(* IEC 61131-3 sources: plcassist-cli/packages/volt-lsp-iec/test-corpus/bakon-nano/Device/Plc Logic/Application/POUs/Calculations (part 2) *)

(* ---- Calc_Hor.fun ---- *)
function Calc_Hor : bool
VAR
	nNrOfLines: INT;
	rLengthOfLine: REAL;
	nNumberOfCutsPerLine: INT;
	nCnt_pos: INT;
	nCnt_line: INT;
	nCnt_Push: INT;
	bToggle: BOOL;
	//nFirstPos: INT;
	//nFirstWastePos: INT;
	rLast_Y_Pos	:REAL;
	rSizeTrimRear	:REAL;
	rSizeTrimFront	:REAL;
	rSizeTrimRight	:REAL;
	rSizeTrimLeft	:REAL;

	//CorrectOvershootHor1a	: CorrectOvershootHor;
	//CorrectOvershootHor1b	: CorrectOvershootHor;
	//CorrectOvershootHor2	: CorrectOvershootHor;
	//CorrectOvershootHor3	: CorrectOvershootHor;
	//CorrectOvershootHor4	: CorrectOvershootHor;
	//CorrectOvershootHor5	: CorrectOvershootHor;
	//CorrectOvershootHor6	: CorrectOvershootHor;
	//CorrectOvershootHor7	: CorrectOvershootHor;
	rMaxTraySize: REAL;
	rMinTraySize: REAL;
	rProdLength_InY: REAL;
	rProdLength_InX: REAL;
	rMmPerCut :REAL;
	rCenterPointKnifeInverted: REAL;
	rSizeOfKnife: REAL;
	//rStartPointTray_Y: REAL;
	rMinimumTrayTrimSize: REAL;
	rNrOfLines 	:REAL;
	rWasteExtra	:REAL;
	rIcedOffset	:REAL;

	rCenterPointKnife: REAL;
	rMinimumSlabTrimSize: REAL;
	nPartsY: INT;

	FirstPoint					: Gonio_Point;
	CopyPoint					: Gonio_Point;

	rFirstYPosition : REAL;
	overshootSettings 			: Gonio_Settings;
	nFirstPosFirstTray 		:INT;
	nFirstWastePosFirstTray :INT;
	nLastPosFirstTray		: INT;
	nLastWastePosFirstTray	: int;
END_VAR

(* Calc_Hor, (mes 0 graden *)

(************************************************************************************************************************************
 * HISTORY
 ************************************************************************************************************************************
 * Update 		: 0.1
 * Author 		: K. Kole
 * Changes	: Tray square, 	calculation for rSizeTrimRight and rSizeTrimLeft changed
 * Update 		: 0.2
 * Author 		: K. Kole
 * Changes	: Tray square, 	calculation for rSizeTrimRear and rSizeTrimFront changed
 ************************************************************************************************************************************)
Calc_Hor := FALSE;
bToggle	:= FALSE;
//nFirstPos := g_sCuttingPositionsInfo.index;
//nFirstWastePos := g_sWastePositionsInfo.index ;

nFirstPosFirstTray 				:= g_sCuttingPositionsInfo.index;
nFirstWastePosFirstTray 		:= g_sWastePositionsInfo.index;

rSizeOfKnife					:= g_HMI_MCH_Parameters.rSizeOfKnife;
rCenterPointKnife				:= rSizeOfKnife/2;
rCenterPointKnifeInverted	:= rSizeOfKnife/2;

overshootSettings.knifeAxis		:= rCenterPointKnife;
overshootSettings.knifeLength	:= rSizeOfKnife;
overshootSettings.precision		:= 0.1;

(**********************************************************************************************************************************)
(* Tray square *)(*AC 23-10-2012 Also Tray Triangle*)
(**********************************************************************************************************************************)
IF		((g_HMI_RCP_Parameters.nProductType = Prod_Tray_Rectangle_1x1)
	OR	(g_HMI_RCP_Parameters.nProductType = Prod_Tray_Rectangle_1x2)
	OR	(g_HMI_RCP_Parameters.nProductType = Prod_Tray_Rectangle_1x4)
	OR 	(g_HMI_RCP_Parameters.nProductType = Prod_Tray_Rectangle_2x1))
THEN

	(* Determine type of tray *)
	IF  (g_HMI_RCP_Parameters.nProductType = Prod_Tray_Rectangle_1x1) THEN
		rProdLength_InY	:= g_HMI_MCH_Parameters.rProdLengthTrayLarge_InY;
		rProdLength_InX	:= g_HMI_MCH_Parameters.rProdLengthTrayLarge_InX;
		rMinimumTrayTrimSize :=	g_HMI_MCH_Parameters.rMinimumTrimSizeTrayLarge;
		FirstPoint.X := g_HMI_MCH_Parameters.rStartPointTrayLarge_X;
		FirstPoint.Y := g_HMI_MCH_Parameters.rStartPointTrayLarge_Y;
	ELSIF	(g_HMI_RCP_Parameters.nProductType = Prod_Tray_Rectangle_1x2)
	THEN
		rProdLength_InY	:= g_HMI_MCH_Parameters.rProdLengthTraySmall_InY;
		rProdLength_InX	:= g_HMI_MCH_Parameters.rProdLengthTraySmall_InX;
		rMinimumTrayTrimSize :=	g_HMI_MCH_Parameters.rMinimumTrimSizeTraySmall;
		FirstPoint.X  := g_HMI_MCH_Parameters.rStartPointTraySmall_X;
		FirstPoint.Y  := g_HMI_MCH_Parameters.rStartPointTraySmall1_Y;	(* Startpoint for first small tray *)
	ELSIF	(g_HMI_RCP_Parameters.nProductType = Prod_Tray_Rectangle_1x4)
	THEN
		rProdLength_InY	:= g_HMI_MCH_Parameters.rProdLengthTrayTriple_InY;
		rProdLength_InX	:= g_HMI_MCH_Parameters.rProdLengthTrayTriple_InX;
		rMinimumTrayTrimSize :=	g_HMI_MCH_Parameters.rMinimumTrimSizeTrayTriple;
		FirstPoint.X  := g_HMI_MCH_Parameters.rStartPointTrayTriple_X;
		FirstPoint.Y  := g_HMI_MCH_Parameters.rStartPointTrayTriple1_Y;	(* Startpoint for first small tray *)
	ELSIF	(g_HMI_RCP_Parameters.nProductType = Prod_Tray_Rectangle_2x1)
	THEN
		rProdLength_InY	:= g_HMI_MCH_Parameters.rProdLengthTrayDouble_InY;
		rProdLength_InX	:= g_HMI_MCH_Parameters.rProdLengthTrayDouble_InX;
		rMinimumTrayTrimSize :=	g_HMI_MCH_Parameters.rMinimumTrimSizeTrayDouble;
		FirstPoint.X  := g_HMI_MCH_Parameters.rStartPointTrayDouble1_X;
		FirstPoint.Y  := g_HMI_MCH_Parameters.rStartPointTrayDouble_Y;	(* Startpoint for first small tray *)
	END_IF

	IF g_HMI_RCP_Parameters.bTrianglesInTray AND g_HMI_RCP_Parameters.bUseRectanglesInEight THEN (*AC 04-07-2013: Uitbreiding 8 driehoeken uit stuk*)
		nPartsY := g_HMI_RCP_Parameters.nPartsY * 2;
	ELSE
		nPartsY := g_HMI_RCP_Parameters.nPartsY;
	END_IF

	IF g_HMI_RCP_Parameters.rSizeTrimFront <= 0			(* Wijziging 16 juli 2010 *)(*AC 28-11-12: Omgedraaid vanaf HMI INstellingen*)
	THEN
		rSizeTrimRear	:= 0;
	ELSE
		rSizeTrimRear 	:= MAX(rMinimumTrayTrimSize, g_HMI_RCP_Parameters.rSizeTrimFront); (*AC 28-11-12: Omgedraaid vanaf HMI INstellingen*)
	END_IF
	IF g_HMI_RCP_Parameters.rSizeTrimRear<= 0			(* Wijziging 16 juli 2010 *)(*AC 28-11-12: Omgedraaid vanaf HMI INstellingen*)
	THEN
		rSizeTrimFront	:= 0;
	ELSE
		rSizeTrimFront 	:= MAX(rMinimumTrayTrimSize, g_HMI_RCP_Parameters.rSizeTrimRear);(*AC 28-11-12: Omgedraaid vanaf HMI INstellingen*)
	END_IF
	rSizeTrimRight 	:= MAX(rMinimumTrayTrimSize, g_HMI_RCP_Parameters.rSizeTrimRight);
	rSizeTrimLeft 		:= MAX(rMinimumTrayTrimSize, g_HMI_RCP_Parameters.rSizeTrimLeft);

	(*Additional safety checks for trays*)
	rMaxTraySize := rProdLength_InX - (rMinimumTrayTrimSize * 2);
	IF			rMaxTraySize >= (g_HMI_MCH_Parameters.rSizeOfKnife)											(* Fixed mes past in het blik *)
	THEN
		rSizeOfKnife					:= g_HMI_MCH_Parameters.rSizeOfKnife;
		rCenterPointKnife				:= rSizeOfKnife/2;
		rCenterPointKnifeInverted	:= rSizeOfKnife/2;
		rMinTraySize					:= rProdLength_InX - (rSizeTrimRight + rSizeTrimLeft);
		IF rMinTraySize < rSizeOfKnife THEN
			rSizeTrimRight	:= rSizeTrimRight - (rSizeOfKnife - rMinTraySize);
			rSizeTrimRight 	:= MAX(rMinimumTrayTrimSize, rSizeTrimRight);								(* Check if new calculated trim is >= MinimumTrim *)
			rSizeTrimLeft	:= rProdLength_InX - rSizeOfKnife - rSizeTrimRight;
		END_IF
	ELSE																											(* Fixed mes past NIET in het blik *)
		g_sMACH.ERR.bTrayTooSmall := TRUE;
		RETURN;
	END_IF

	g_rDistanceBetweenCuts_InY:=	(rProdLength_InY - rSizeTrimRear - rSizeTrimFront) / INT_TO_REAL(nPartsY);(*g_HMI_RCP_Parameters.nPartsY);*)

	(* Determine number of lines *)
	IF g_bTrimRear AND g_bTrimFront
	THEN
		nNrOfLines	:= 1 + nPartsY;(*g_HMI_RCP_Parameters.nPartsY);*)(*AC 04-07-2013*)
	ELSIF g_bTrimRear AND NOT g_bTrimFront
	THEN
		nNrOfLines	:= nPartsY;(*g_HMI_RCP_Parameters.nPartsY);*)(*AC 04-07-2013*)
	ELSIF NOT g_bTrimRear AND g_bTrimFront
	THEN
		nNrOfLines	:= nPartsY;(*g_HMI_RCP_Parameters.nPartsY);*)(*AC 04-07-2013*)
	ELSIF NOT g_bTrimRear AND NOT g_bTrimFront
	THEN
		nNrOfLines	:=nPartsY - 1;(*g_HMI_RCP_Parameters.nPartsY);*)(*AC 04-07-2013*)
	END_IF

	(* Calculate number of cuts on the line *)
	rLengthOfLine := rProdLength_InX - rSizeTrimRight - rSizeTrimLeft;
	IF rLengthOfLine > rSizeOfKnife
	THEN
		nNumberOfCutsPerLine := TRUNC_INT(rLengthOfLine / rSizeOfKnife);
		IF nNumberOfCutsPerLine < (rLengthOfLine / rSizeOfKnife)
		THEN
			nNumberOfCutsPerLine := nNumberOfCutsPerLine + 1;
		END_IF
	ELSE
		nNumberOfCutsPerLine := 1;
	END_IF
	(*Calculation of covered distance per cut*)
	rMmPerCut := (rLengthOfLine - rSizeOfKnife)/(nNumberOfCutsPerLine -1);

	(* Calculate positions on first line *)
	overshootSettings.MarginXMin := FirstPoint.x + MAX(rMinimumTrayTrimSize-0.1,1);		(* Mechanical boundary *)
	overshootSettings.MarginXMax := FirstPoint.x + rProdLength_InX  - MAX(rMinimumTrayTrimSize-0.1,1);	(* Mechanical boundary *)
	overshootSettings.MarginYMin := FirstPoint.y + MAX(rMinimumTrayTrimSize-0.1,1);		(* Mechanical boundary *)
	overshootSettings.MarginYMax := FirstPoint.y + rProdLength_InY -  MAX(rMinimumTrayTrimSize-0.1,1);		(* Mechanical boundary *)

	overshootSettings.adjustXMax := FALSE;
	overshootSettings.adjustXMin := FALSE;
	overshootSettings.adjustYMax := FALSE;
	overshootSettings.adjustYMin := FALSE;

	IF g_bTrimRear
	THEN
		IF nNumberOfCutsPerLine = 1
		THEN
			IF NOT StorePos(I_rX:= 							Firstpoint.X + rSizeTrimRight + rCenterPointKnife,
							I_rY:=							(rFirstYPosition := Firstpoint.Y + rSizeTrimRear),
							I_rA:=							0,
							I_rK:=							0,
							I_bIsWaste :=					 (g_HMI_RCP_Parameters.bCutWasteFirst) ,
							I_sOvershootSettings := 		overshootSettings)
			THEN
								RETURN;
			END_IF
		ELSE
			FOR nCnt_pos:=1 TO (nNumberOfCutsPerLine - 1) DO
				IF NOT StorePos(I_rX:= 							FirstPoint.X + rSizeTrimRight + (nCnt_pos - 1) * rMmPerCut
																			 + rCenterPointKnife,
								I_rY:=							(rFirstYPosition := FirstPoint.Y + rSizeTrimRear),
								I_rA:=							0,
								I_rK:=							0,
								I_bIsWaste :=					 (g_HMI_RCP_Parameters.bCutWasteFirst) ,
								I_sOvershootSettings := 		overshootSettings)
				THEN
										RETURN;
				END_IF
			END_FOR
			(* Last position on the line *)
			IF NOT StorePos(I_rX:= 							Firstpoint.X + rProdLength_InX - rSizeTrimLeft - rCenterPointKnifeInverted,
							I_rY:=							Firstpoint.Y + rSizeTrimRear,
							I_rA:=							0,
							I_rK:=							0,
							I_bIsWaste :=					 (g_HMI_RCP_Parameters.bCutWasteFirst) ,
							I_sOvershootSettings := 		overshootSettings)
			THEN
								RETURN;
			END_IF

		END_IF
	ELSE (* No waste strip at the left *)
		IF nNrOfLines > 0	(* New 8 feb 2010: when only one piece and no trims *)
		THEN
			IF nNumberOfCutsPerLine = 1
			THEN
				IF NOT StorePos(I_rX:= 							Firstpoint.X + rSizeTrimRight + rCenterPointKnife,
								I_rY:=							(rFirstYPosition := Firstpoint.Y + rSizeTrimRear + g_rDistanceBetweenCuts_InY),
								I_rA:=							0,
								I_rK:=							0,
								I_bIsWaste :=					FALSE,
								I_sOvershootSettings := 		overshootSettings)
				THEN
										RETURN;
				END_IF

			ELSE
				FOR nCnt_pos:=1 TO (nNumberOfCutsPerLine - 1) DO
					IF NOT StorePos(I_rX:= 							Firstpoint.X + rSizeTrimRight + (nCnt_pos - 1) * rMmPerCut
																					 + rCenterPointKnife,
									I_rY:=							(rFirstYPosition := Firstpoint.Y + rSizeTrimRear + g_rDistanceBetweenCuts_InY),
									I_rA:=							0,
									I_rK:=							0,
									I_bIsWaste :=					FALSE,
									I_sOvershootSettings := 		overshootSettings)
					THEN
												RETURN;
					END_IF

				END_FOR
				(* Last position on the line *)
				IF NOT StorePos(I_rX:= 							Firstpoint.X + rProdLength_InX - rSizeTrimLeft - rCenterPointKnifeInverted,
								I_rY:=							Firstpoint.Y + rSizeTrimRear + g_rDistanceBetweenCuts_InY,
								I_rA:=							0,
								I_rK:=							0,
								I_bIsWaste :=					FALSE,
								I_sOvershootSettings := 		overshootSettings)
				THEN
										RETURN;
				END_IF

			END_IF
		END_IF
	END_IF

	(* Fill in all other positions on the rest of the lines *)

	FOR nCnt_line := 2 TO (nNrOfLines) BY 1 DO
		IF nNumberOfCutsPerLine = 1
		THEN
			IF NOT StorePos(I_rX:= 							Firstpoint.X + rSizeTrimRight + rCenterPointKnife,
							I_rY:=							rFirstYPosition + (nCnt_line-1) * g_rDistanceBetweenCuts_InY,
							I_rA:=							0,
							I_rK:=							0,
							I_bIsWaste :=					 (g_HMI_RCP_Parameters.bCutWasteFirst AND g_bTrimFront AND nCnt_Line = nNrOfLines) ,
							I_sOvershootSettings := 		overshootSettings)
			THEN
								RETURN;
			END_IF

		ELSE
			IF bToggle (* from front to rear *)
			THEN
				FOR nCnt_pos:=1 TO (nNumberOfCutsPerLine - 1) DO
					IF NOT StorePos(I_rX:= 							Firstpoint.X + rSizeTrimRight + rCenterPointKnife
														                                                   + (nCnt_pos - 1) * rMmPerCut ,
									I_rY:=							rFirstYPosition + (nCnt_line-1) * g_rDistanceBetweenCuts_InY,
									I_rA:=							0,
									I_rK:=							0,
									I_bIsWaste :=					 (g_HMI_RCP_Parameters.bCutWasteFirst AND g_bTrimFront AND nCnt_Line = nNrOfLines) ,
									I_sOvershootSettings := 		overshootSettings)
					THEN
												RETURN;
					END_IF

				END_FOR
				(* Last position on the line *)
				IF NOT StorePos(I_rX:= 							Firstpoint.X + rProdLength_InX - rSizeTrimLeft - rCenterPointKnifeInverted,
								I_rY:=							rFirstYPosition + (nCnt_line-1) * g_rDistanceBetweenCuts_InY,
								I_rA:=							0,
								I_rK:=							0,
								I_bIsWaste :=					 (g_HMI_RCP_Parameters.bCutWasteFirst AND g_bTrimFront AND nCnt_Line = nNrOfLines) ,
								I_sOvershootSettings := 		overshootSettings)
				THEN
										RETURN;
				END_IF

			ELSE (* toggle, ie from rear to front *)
				FOR nCnt_pos:=1 TO (nNumberOfCutsPerLine - 1) DO
					IF NOT StorePos(I_rX:= 							Firstpoint.X + rProdLength_InX - rSizeTrimLeft - rCenterPointKnifeInverted
																					- (nCnt_pos -1) * rMmPerCut,
									I_rY:=							rFirstYPosition + (nCnt_line-1) * g_rDistanceBetweenCuts_InY,
									I_rA:=							0,
									I_rK:=							0,
									I_bIsWaste :=					 (g_HMI_RCP_Parameters.bCutWasteFirst AND g_bTrimFront AND nCnt_Line = nNrOfLines) ,
									I_sOvershootSettings := 		overshootSettings)
					THEN
												RETURN;
					END_IF

				END_FOR
				(* Last position on the line *)
				IF NOT StorePos(I_rX:= 							FirstPoint.X + rSizeTrimRight + rCenterPointKnife,
								I_rY:=							rFirstYPosition + (nCnt_line-1) * g_rDistanceBetweenCuts_InY,
								I_rA:=							0,
								I_rK:=							0,
								I_bIsWaste :=					 (g_HMI_RCP_Parameters.bCutWasteFirst AND g_bTrimFront AND nCnt_Line = nNrOfLines) ,
								I_sOvershootSettings := 		overshootSettings)
				THEN
										RETURN;
				END_IF

			END_IF
			bToggle := NOT bToggle;
		END_IF
	END_FOR

	nLastPosFirstTray		:= g_sCuttingPositionsInfo.index-1;
	nLastWastePosFirstTray	:= g_sWastePositionsInfo.index-1;

	(* Double the positions for the second tray if small trays is selected *)
	IF	g_HMI_RCP_Parameters.nProductType = Prod_Tray_Rectangle_1x2
	THEN

		CopyPoint.X := FirstPoint.X;
		CopyPoint.Y := g_HMI_MCH_Parameters.rStartPointTraySmall2_Y;

		overshootSettings.MarginXMin := CopyPoint.X + MAX(rMinimumTrayTrimSize-0.1,1);		(* Mechanical boundary *)
		overshootSettings.MarginXMax := CopyPoint.X + rProdLength_InX  - MAX(rMinimumTrayTrimSize-0.1,1);	(* Mechanical boundary *)
		overshootSettings.MarginYMin := CopyPoint.Y + MAX(rMinimumTrayTrimSize-0.1,1);		(* Mechanical boundary *)
		overshootSettings.MarginYMax := CopyPoint.Y + rProdLength_InY -  MAX(rMinimumTrayTrimSize-0.1,1);		(* Mechanical boundary *)

		IF nFirstPosFirstTray <= nLastPosFirstTray THEN
			IF NOT Calc_CopyCutsWithOffset(
				I_firstIndex				:= nFirstPosFirstTray,
				I_lastIndex					:= nLastPosFirstTray,
				I_dX 						:= CopyPoint.X - FirstPoint.X,
				I_dY 						:= CopyPoint.Y - FirstPoint.Y,
				I_overshootSettings 		:= overshootSettings,
				I_dataArray 				:= ADR(g_aCuttingPositions),
				I_bReverseOrder				:= (nNrOfLines MOD 2)>0,
				IQ_dataArrayInfo 			:= g_sCuttingPositionsInfo)
			THEN
								RETURN;
			END_IF
		END_IF

		IF nFirstWastePosFirstTray <= nLastWastePosFirstTray THEN
			IF NOT Calc_CopyCutsWithOffset(
				I_firstIndex				:= nFirstWastePosFirstTray,
				I_lastIndex					:= nLastWastePosFirstTray,
				I_dX 						:= CopyPoint.X - FirstPoint.X,
				I_dY 						:= CopyPoint.Y - FirstPoint.Y,
				I_overshootSettings 		:= overshootSettings,
				I_dataArray 				:= ADR(g_aWastePositions),
				I_bReverseOrder				:= (nNrOfLines MOD 2)>0,
				IQ_dataArrayInfo 			:= g_sWastePositionsInfo)
			THEN
								RETURN;
			END_IF
		END_IF
	END_IF

	(* Triple the positions for the second and third tray if triple trays is selected *)
	IF	g_HMI_RCP_Parameters.nProductType = Prod_Tray_Rectangle_1x4
	THEN

		CopyPoint.X := FirstPoint.X;
		CopyPoint.Y := g_HMI_MCH_Parameters.rStartPointTrayTriple2_Y;

		overshootSettings.MarginXMin := CopyPoint.X + MAX(rMinimumTrayTrimSize-0.1,1);		(* Mechanical boundary *)
		overshootSettings.MarginXMax := CopyPoint.X + rProdLength_InX  - MAX(rMinimumTrayTrimSize-0.1,1);	(* Mechanical boundary *)
		overshootSettings.MarginYMin := CopyPoint.Y + MAX(rMinimumTrayTrimSize-0.1,1);		(* Mechanical boundary *)
		overshootSettings.MarginYMax := CopyPoint.Y + rProdLength_InY -  MAX(rMinimumTrayTrimSize-0.1,1);		(* Mechanical boundary *)

		IF nFirstPosFirstTray <= nLastPosFirstTray THEN
			IF NOT Calc_CopyCutsWithOffset(
				I_firstIndex				:= nFirstPosFirstTray,
				I_lastIndex					:= nLastPosFirstTray,
				I_dX 						:= CopyPoint.X - FirstPoint.X,
				I_dY 						:= CopyPoint.Y - FirstPoint.Y,
				I_overshootSettings 		:= overshootSettings,
				I_dataArray 				:= ADR(g_aCuttingPositions),
				I_bReverseOrder				:= (nNrOfLines MOD 2)>0,
				IQ_dataArrayInfo 			:= g_sCuttingPositionsInfo)
			THEN
								RETURN;
			END_IF
		END_IF

		IF nFirstWastePosFirstTray <= nLastWastePosFirstTray THEN
			IF NOT Calc_CopyCutsWithOffset(
				I_firstIndex				:= nFirstWastePosFirstTray,
				I_lastIndex					:= nLastWastePosFirstTray,
				I_dX 						:= CopyPoint.X - FirstPoint.X,
				I_dY 						:= CopyPoint.Y - FirstPoint.Y,
				I_overshootSettings 		:= overshootSettings,
				I_dataArray 				:= ADR(g_aWastePositions),
				I_bReverseOrder				:= (nNrOfLines MOD 2)>0,
				IQ_dataArrayInfo 			:= g_sWastePositionsInfo)
			THEN
								RETURN;
			END_IF
		END_IF

		(*Third tray*)
		CopyPoint.X := FirstPoint.X;
		CopyPoint.Y := g_HMI_MCH_Parameters.rStartPointTrayTriple3_Y;

		overshootSettings.MarginXMin := CopyPoint.X + MAX(rMinimumTrayTrimSize-0.1,1);		(* Mechanical boundary *)
		overshootSettings.MarginXMax := CopyPoint.X + rProdLength_InX  - MAX(rMinimumTrayTrimSize-0.1,1);	(* Mechanical boundary *)
		overshootSettings.MarginYMin := CopyPoint.Y + MAX(rMinimumTrayTrimSize-0.1,1);		(* Mechanical boundary *)
		overshootSettings.MarginYMax := CopyPoint.Y + rProdLength_InY -  MAX(rMinimumTrayTrimSize-0.1,1);		(* Mechanical boundary *)

		IF nFirstPosFirstTray <= nLastPosFirstTray THEN
			IF NOT Calc_CopyCutsWithOffset(
				I_firstIndex				:= nFirstPosFirstTray,
				I_lastIndex					:= nLastPosFirstTray,
				I_dX 						:= CopyPoint.X - FirstPoint.X,
				I_dY 						:= CopyPoint.Y - FirstPoint.Y,
				I_overshootSettings 		:= overshootSettings,
				I_dataArray 				:= ADR(g_aCuttingPositions),
				I_bReverseOrder				:= FALSE,
				IQ_dataArrayInfo 			:= g_sCuttingPositionsInfo)
			THEN
								RETURN;
			END_IF
		END_IF

		IF nFirstWastePosFirstTray <= nLastWastePosFirstTray THEN
			IF NOT Calc_CopyCutsWithOffset(
				I_firstIndex				:= nFirstWastePosFirstTray,
				I_lastIndex					:= nLastWastePosFirstTray,
				I_dX 						:= CopyPoint.X - FirstPoint.X,
				I_dY 						:= CopyPoint.Y - FirstPoint.Y,
				I_overshootSettings 		:= overshootSettings,
				I_dataArray 				:= ADR(g_aWastePositions),
				I_bReverseOrder				:= FALSE,
				IQ_dataArrayInfo 			:= g_sWastePositionsInfo)
			THEN
								RETURN;
			END_IF
		END_IF

		(*Fourth Tray*)
		CopyPoint.X := FirstPoint.X;
		CopyPoint.Y := g_HMI_MCH_Parameters.rStartPointTrayTriple4_Y;

		overshootSettings.MarginXMin := CopyPoint.X + MAX(rMinimumTrayTrimSize-0.1,1);		(* Mechanical boundary *)
		overshootSettings.MarginXMax := CopyPoint.X + rProdLength_InX  - MAX(rMinimumTrayTrimSize-0.1,1);	(* Mechanical boundary *)
		overshootSettings.MarginYMin := CopyPoint.Y + MAX(rMinimumTrayTrimSize-0.1,1);		(* Mechanical boundary *)
		overshootSettings.MarginYMax := CopyPoint.Y + rProdLength_InY -  MAX(rMinimumTrayTrimSize-0.1,1);		(* Mechanical boundary *)

		IF nFirstPosFirstTray <= nLastPosFirstTray THEN
			IF NOT Calc_CopyCutsWithOffset(
				I_firstIndex				:= nFirstPosFirstTray,
				I_lastIndex					:= nLastPosFirstTray,
				I_dX 						:= CopyPoint.X - FirstPoint.X,
				I_dY 						:= CopyPoint.Y - FirstPoint.Y,
				I_overshootSettings 		:= overshootSettings,
				I_dataArray 				:= ADR(g_aCuttingPositions),
				I_bReverseOrder				:= (nNrOfLines MOD 2)>0,
				IQ_dataArrayInfo 			:= g_sCuttingPositionsInfo)
			THEN
								RETURN;
			END_IF
		END_IF

		IF nFirstWastePosFirstTray <= nLastWastePosFirstTray THEN
			IF NOT Calc_CopyCutsWithOffset(
				I_firstIndex				:= nFirstWastePosFirstTray,
				I_lastIndex					:= nLastWastePosFirstTray,
				I_dX 						:= CopyPoint.X - FirstPoint.X,
				I_dY 						:= CopyPoint.Y - FirstPoint.Y,
				I_overshootSettings 		:= overshootSettings,
				I_dataArray 				:= ADR(g_aWastePositions),
				I_bReverseOrder				:= (nNrOfLines MOD 2)>0,
				IQ_dataArrayInfo 			:= g_sWastePositionsInfo)
			THEN
								RETURN;
			END_IF
		END_IF
	END_IF

	(* 2x positions the positions for the second tray if double trays side by side *)
	IF	g_HMI_RCP_Parameters.nProductType = Prod_Tray_Rectangle_2x1
	THEN
		CopyPoint.X := g_HMI_MCH_Parameters.rStartPointTrayDouble2_X; // FirstPoint.X;
		CopyPoint.Y := FirstPoint.Y;// g_HMI_MCH_Parameters.rStartPointTrayDouble2_X;

		overshootSettings.MarginXMin := CopyPoint.X + MAX(rMinimumTrayTrimSize-0.1,1);		(* Mechanical boundary *)
		overshootSettings.MarginXMax := CopyPoint.X + rProdLength_InX  - MAX(rMinimumTrayTrimSize-0.1,1);	(* Mechanical boundary *)
		overshootSettings.MarginYMin := CopyPoint.Y + MAX(rMinimumTrayTrimSize-0.1,1);		(* Mechanical boundary *)
		overshootSettings.MarginYMax := CopyPoint.Y + rProdLength_InY -  MAX(rMinimumTrayTrimSize-0.1,1);		(* Mechanical boundary *)

		IF nFirstPosFirstTray <= nLastPosFirstTray THEN
			IF NOT Calc_CopyCutsWithOffset(
				I_firstIndex				:= nFirstPosFirstTray,
				I_lastIndex					:= nLastPosFirstTray,
				I_dX 						:= CopyPoint.X - FirstPoint.X,
				I_dY 						:= CopyPoint.Y - FirstPoint.Y,
				I_overshootSettings 		:= overshootSettings,
				I_dataArray 				:= ADR(g_aCuttingPositions),
				I_bReverseOrder				:= true,
				IQ_dataArrayInfo 			:= g_sCuttingPositionsInfo)
			THEN
								RETURN;
			END_IF
		END_IF

		IF nFirstWastePosFirstTray <= nLastWastePosFirstTray THEN
			IF NOT Calc_CopyCutsWithOffset(
				I_firstIndex				:= nFirstWastePosFirstTray,
				I_lastIndex					:= nLastWastePosFirstTray,
				I_dX 						:= CopyPoint.X - FirstPoint.X,
				I_dY 						:= CopyPoint.Y - FirstPoint.Y,
				I_overshootSettings 		:= overshootSettings,
				I_dataArray 				:= ADR(g_aWastePositions),
				I_bReverseOrder				:= true,
				IQ_dataArrayInfo 			:= g_sWastePositionsInfo)
			THEN
								RETURN;
			END_IF
		END_IF
	END_IF

(**********************************************************************************************************************************)
(* If slab (square or diagonal) *)
(**********************************************************************************************************************************)
ELSIF 		(g_HMI_RCP_Parameters.nProductType = Prod_Slab_Rectangle_1x1)
		OR	(g_HMI_RCP_Parameters.nProductType = Prod_Slab_Diagonal_1x1)
		OR	(g_HMI_RCP_Parameters.nProductType = Prod_Slab_Rectangle_1x1_Clamp)		(* V04.01 *)
THEN
	IF g_HMI_RCP_Parameters.nProductType = Prod_Slab_Rectangle_1x1 THEN
		rIcedOffset 				:= g_HMI_RCP_Parameters.rShiftCompensation;
		rMinimumSlabTrimSize	:= 0;
	ELSE
		rIcedOffset := 0;
		IF	(g_HMI_RCP_Parameters.nProductType = Prod_Slab_Rectangle_1x1_Clamp) THEN
			rIcedOffset 				:= g_HMI_RCP_Parameters.rShiftCompensation;
			rMinimumSlabTrimSize	:= g_HMI_MCH_Parameters.rMinimumTrimSizeSlab;
		ELSE
			rMinimumSlabTrimSize	:= 0;
		END_IF
	END_IF

	rSizeOfKnife					:= g_HMI_MCH_Parameters.rSizeOfKnife;
	rCenterPointKnife				:= rSizeOfKnife/2;
	rCenterPointKnifeInverted	:= rSizeOfKnife/2;

	(* Offset of slab *)
	FirstPoint.X	:= g_HMI_MCH_Parameters.rStartPointSlab_X;
	FirstPoint.Y	:= g_HMI_MCH_Parameters.rStartPointSlab_Y;

	rProdLength_InX	:= g_HMI_RCP_Parameters.rProdLength_InX + (rIcedOffset * g_HMI_RCP_Parameters.nPartsX);
	rProdLength_InY 	:= g_HMI_RCP_Parameters.rProdLength_InY;

	IF	(g_HMI_RCP_Parameters.nProductType = Prod_Slab_Rectangle_1x1_Clamp)		(* V04.01 *)
	THEN
		IF g_HMI_RCP_Parameters.rSizeTrimFront <= 0
		THEN
			rSizeTrimRear 	:= 0;
			//rSizeTrimRear 	:= MAX(rMinimumSlabTrimSize, g_HMI_RCP_Parameters.rSizeTrimFront); sept 2016
		ELSE
			rSizeTrimRear 	:= MAX(rMinimumSlabTrimSize, g_HMI_RCP_Parameters.rSizeTrimFront);
		END_IF
		IF g_HMI_RCP_Parameters.rSizeTrimRear<= 0			(* Omgedraaid vanaf HMI Instellingen*)
		THEN
			rSizeTrimFront	:= 0;
		ELSE
			rSizeTrimFront 	:= MAX(0, g_HMI_RCP_Parameters.rSizeTrimRear);(*Omgedraaid vanaf HMI INstellingen*)
		END_IF
		rSizeTrimRight 	:= MAX(rMinimumSlabTrimSize, g_HMI_RCP_Parameters.rSizeTrimRight);
		rSizeTrimLeft 	:= MAX(rMinimumSlabTrimSize, g_HMI_RCP_Parameters.rSizeTrimLeft);
		//rSizeTrimLeft 		:= MAX(0, g_HMI_RCP_Parameters.rSizeTrimLeft); sept 2016

		(*Additional safety checks for slab with fingers *)
		(*rMaxSlabSize := rProdLength_InX - (rMinimumSlabTrimSize);
		IF			rMaxSlabSize >= (g_HMI_MCH_Parameters.rSizeOfKnife)											(* Fixed mes past in de slab tussen de vingers *)
		THEN
			rMinSlabSize					:= rProdLength_InX - (rSizeTrimRight + rSizeTrimLeft);
			IF rMinSlabSize < rSizeOfKnife THEN
				rSizeTrimRight	:= rSizeTrimRight - (rSizeOfKnife - rMinSlabSize);
				rSizeTrimRight 	:= MAX(rMinimumSlabTrimSize, rSizeTrimRight);								(* Check if new calculated trim is >= MinimumTrim *)
				rSizeTrimLeft		:= rProdLength_InX - rSizeOfKnife - rSizeTrimRight;
			END_IF
		ELSE																											(* Fixed mes past NIET in het blik *)
			g_sMACH.ERR.bSlabTooSmall := TRUE;
			RETURN;
		END_IF*)
	ELSE
		rSizeTrimRear 	:= MAX(0, g_HMI_RCP_Parameters.rSizeTrimFront);(*AC 28-11-12: Omgedraaid vanaf HMI INstellingen*)
		rSizeTrimFront 	:= MAX(0, g_HMI_RCP_Parameters.rSizeTrimRear); (*AC 28-11-12: Omgedraaid vanaf HMI INstellingen*)
		rSizeTrimRight 	:= g_HMI_RCP_Parameters.rSizeTrimRight;
		rSizeTrimLeft 	:= g_HMI_RCP_Parameters.rSizeTrimLeft;
	END_IF

	g_rDistanceBetweenCuts_InY:=	(rProdLength_InY - rSizeTrimRear - rSizeTrimFront) / INT_TO_REAL(g_HMI_RCP_Parameters.nPartsY);

	(* Determine number of lines *)
	IF g_bTrimRear AND g_bTrimFront
	THEN
		nNrOfLines	:= g_HMI_RCP_Parameters.nPartsY + 1;
	ELSIF g_bTrimRear AND NOT g_bTrimFront
	THEN
		nNrOfLines	:= g_HMI_RCP_Parameters.nPartsY;
	ELSIF NOT g_bTrimRear AND g_bTrimFront
	THEN
		nNrOfLines	:= g_HMI_RCP_Parameters.nPartsY;
	ELSIF NOT g_bTrimRear AND NOT g_bTrimFront
	THEN
		nNrOfLines	:= g_HMI_RCP_Parameters.nPartsY - 1;
	END_IF

	IF	(g_HMI_RCP_Parameters.nProductType = Prod_Slab_Rectangle_1x1_Clamp)		(* V04.01 *)
	THEN
		overshootSettings.MarginXMin := FirstPoint.X + rSizeTrimRight;
		overshootSettings.MarginXMax := SEL(gMachConfig.bXL,C_rMaxOvershootX,C_rMaxOvershootX_XL);
		overshootSettings.MarginYMin := FirstPoint.Y + rSizeTrimRear;
		overshootSettings.MarginYMax := SEL(gMachConfig.bXL,C_rMaxOvershootY,C_rMaxOvershootY_XL);
	ELSE
		overshootSettings.MarginXMin := C_rMinOvershootX;
		overshootSettings.MarginXMax := SEL(gMachConfig.bXL,C_rMaxOvershootX,C_rMaxOvershootX_XL);
		overshootSettings.MarginYMin := C_rMinOvershootY;
		overshootSettings.MarginYMax := SEL(gMachConfig.bXL,C_rMaxOvershootY,C_rMaxOvershootY_XL);
	END_IF

	overshootSettings.adjustXMax := TRUE;
	overshootSettings.adjustXMin := NOT (g_HMI_RCP_Parameters.nProductType = Prod_Slab_Rectangle_1x1_Clamp);
	overshootSettings.adjustYMax := TRUE;
	overshootSettings.adjustYMin := NOT (g_HMI_RCP_Parameters.nProductType = Prod_Slab_Rectangle_1x1_Clamp);

	IF nNrOfLines > 0 THEN
		(* Calculate number of cuts on the line *)
		(*rLengthOfLine := g_HMI_RCP_Parameters.rProdLength_InX - rSizeTrimRight - rSizeTrimLeft;*)
		rLengthOfLine := g_HMI_RCP_Parameters.rProdLength_InX - rSizeTrimRight - rSizeTrimLeft + (g_HMI_RCP_Parameters.nPartsX * rIcedOffset); (*AC 28-11-12: Deze richting wordt als tweede gesneden en de plak langer geworden.*)
		IF rLengthOfLine > rSizeOfKnife
		THEN
			nNumberOfCutsPerLine := TRUNC_INT(rLengthOfLine / rSizeOfKnife);
			IF nNumberOfCutsPerLine < (rLengthOfLine / rSizeOfKnife)
			THEN
				nNumberOfCutsPerLine := nNumberOfCutsPerLine + 1;
			END_IF
			rMmPerCut := (rLengthOfLine - rSizeOfKnife)/(nNumberOfCutsPerLine -1);
		ELSE
			nNumberOfCutsPerLine := 1;
		END_IF

		(* Calculate positions on first line *)
		IF g_bTrimRear
		THEN
			IF nNumberOfCutsPerLine = 1
			THEN
				IF NOT StorePos(I_rX:= 							FirstPoint.X + rSizeTrimRight + rCenterPointKnife,
								I_rY:=							(rFirstYPosition := FirstPoint.Y + rSizeTrimRear),
								I_rA:=							0,
								I_rK:=							0,
								I_bIsWaste :=					 (g_HMI_RCP_Parameters.bCutWasteFirst) ,
								I_sOvershootSettings := 		overshootSettings)
				THEN
										RETURN;
				END_IF

			ELSE
				FOR nCnt_pos:=1 TO (nNumberOfCutsPerLine - 1) DO
					IF NOT StorePos(I_rX:= 							FirstPoint.X + rSizeTrimRight + (nCnt_pos - 1) * rMmPerCut
																					 + rCenterPointKnife,
									I_rY:=							(rFirstYPosition := FirstPoint.Y + rSizeTrimRear),
									I_rA:=							0,
									I_rK:=							0,
									I_bIsWaste :=					 (g_HMI_RCP_Parameters.bCutWasteFirst) ,
									I_sOvershootSettings := 		overshootSettings)
					THEN
												RETURN;
					END_IF

				END_FOR
				(* Last position on the line *)
				IF NOT StorePos(I_rX:= 							FirstPoint.X + rProdLength_InX - rSizeTrimLeft - rCenterPointKnifeInverted,
								I_rY:=							FirstPoint.Y + rSizeTrimRear,
								I_rA:=							0,
								I_rK:=							0,
								I_bIsWaste :=					 (g_HMI_RCP_Parameters.bCutWasteFirst) ,
								I_sOvershootSettings := 		overshootSettings)
				THEN
										RETURN;
				END_IF

			END_IF
		ELSE (* No waste strip at the left *)
			IF nNumberOfCutsPerLine = 1
			THEN
				IF NOT StorePos(I_rX:= 							FirstPoint.X + rSizeTrimRight + rCenterPointKnife,
								I_rY:=							(rFirstYPosition := FirstPoint.Y + rSizeTrimRear + g_rDistanceBetweenCuts_InY),
								I_rA:=							0,
								I_rK:=							0,
								I_bIsWaste :=					FALSE,
								I_sOvershootSettings := 		overshootSettings)
				THEN
										RETURN;
				END_IF

			ELSE
				FOR nCnt_pos:=1 TO (nNumberOfCutsPerLine - 1) DO
					IF NOT StorePos(I_rX:= 							FirstPoint.X + rSizeTrimRight + (nCnt_pos - 1) * rMmPerCut
																					 + rCenterPointKnife,
									I_rY:=							(rFirstYPosition := FirstPoint.Y + rSizeTrimRear + g_rDistanceBetweenCuts_InY),
									I_rA:=							0,
									I_rK:=							0,
									I_bIsWaste :=					FALSE,
									I_sOvershootSettings := 		overshootSettings)
					THEN
												RETURN;
					END_IF

				END_FOR
				(* Last position on the line *)
				IF NOT StorePos(I_rX:= 							FirstPoint.X + rProdLength_InX - rSizeTrimLeft - rCenterPointKnifeInverted,
								I_rY:=							FirstPoint.Y + rSizeTrimRear + g_rDistanceBetweenCuts_InY,
								I_rA:=							0,
								I_rK:=							0,
								I_bIsWaste :=					FALSE,
								I_sOvershootSettings := 		overshootSettings)
				THEN
										RETURN;
				END_IF

			END_IF
		END_IF

		(* Fill in all other positions on the rest of the lines *)

		FOR nCnt_line := 2 TO (nNrOfLines) BY 1 DO
			IF nNumberOfCutsPerLine = 1
			THEN
				IF NOT StorePos(I_rX:= 							FirstPoint.X + rSizeTrimRight + rCenterPointKnife,
								I_rY:=							rFirstYPosition + (nCnt_line-1) * (g_rDistanceBetweenCuts_InY + rIcedOffset),
								I_rA:=							0,
								I_rK:=							0,
								I_bIsWaste :=					 (g_HMI_RCP_Parameters.bCutWasteFirst AND g_bTrimFront AND nCnt_Line = nNrOfLines) ,
								I_sOvershootSettings := 		overshootSettings)
				THEN
										RETURN;
				END_IF

			ELSE
				IF bToggle (* from front to rear *)
				THEN
					FOR nCnt_pos:=1 TO (nNumberOfCutsPerLine - 1) DO
						IF NOT StorePos(I_rX:= 							FirstPoint.X + rSizeTrimRight + rCenterPointKnife
																                                                   + (nCnt_pos - 1) * rMmPerCut ,
										I_rY:=							rFirstYPosition + (nCnt_line-1) * (g_rDistanceBetweenCuts_InY + rIcedOffset),
										I_rA:=							0,
										I_rK:=							0,
										I_bIsWaste :=					 (g_HMI_RCP_Parameters.bCutWasteFirst AND g_bTrimFront AND nCnt_Line = nNrOfLines) ,
										I_sOvershootSettings := 		overshootSettings)
						THEN
														RETURN;
						END_IF

					END_FOR
					(* Last position on the line *)
					IF NOT StorePos(I_rX:= 							FirstPoint.X + rProdLength_InX - rSizeTrimLeft - rCenterPointKnifeInverted,
									I_rY:=							rFirstYPosition + (nCnt_line-1) * (g_rDistanceBetweenCuts_InY + rIcedOffset),
									I_rA:=							0,
									I_rK:=							0,
									I_bIsWaste :=					 (g_HMI_RCP_Parameters.bCutWasteFirst AND g_bTrimFront AND nCnt_Line = nNrOfLines) ,
									I_sOvershootSettings := 		overshootSettings)
					THEN
												RETURN;
					END_IF

				ELSE (* toggle, ie from rear to front *)
					FOR nCnt_pos:=1 TO (nNumberOfCutsPerLine - 1) DO
						IF NOT StorePos(I_rX:= 							FirstPoint.X + rProdLength_InX - rSizeTrimLeft - rCenterPointKnifeInverted
																							- (nCnt_pos -1) * rMmPerCut,
										I_rY:=							rFirstYPosition + (nCnt_line-1) * (g_rDistanceBetweenCuts_InY + rIcedOffset),
										I_rA:=							0,
										I_rK:=							0,
										I_bIsWaste :=					 (g_HMI_RCP_Parameters.bCutWasteFirst AND g_bTrimFront AND nCnt_Line = nNrOfLines) ,
										I_sOvershootSettings := 		overshootSettings)
						THEN
														RETURN;
						END_IF

					END_FOR
					(* Last position on the line *)
					IF NOT StorePos(I_rX:= 							FirstPoint.X + rSizeTrimRight + rCenterPointKnife,
									I_rY:=							rFirstYPosition + (nCnt_line-1) * (g_rDistanceBetweenCuts_InY + rIcedOffset),
									I_rA:=							0,
									I_rK:=							0,
									I_bIsWaste :=					 (g_HMI_RCP_Parameters.bCutWasteFirst AND g_bTrimFront AND nCnt_Line = nNrOfLines) ,
									I_sOvershootSettings := 		overshootSettings)
					THEN
												RETURN;
					END_IF

				END_IF
				bToggle := NOT bToggle;
			END_IF
		END_FOR

		(* Schuiven Uitbreiding AC *)
		(*Alle ingevulde posities controleren of Y gelijk is aan uiterste Y*)
		(*Indien ja: set bPushAwayProduct en corresponderende distance.*)
		IF g_bTrimFront THEN
			rLast_Y_Pos := rFirstYPosition + (nNrOfLines-1) * g_rDistanceBetweenCuts_InY;

			FOR nCnt_Push := nFirstPosFirstTray TO g_sCuttingPositionsInfo.index -1 DO
				IF rLast_Y_Pos = g_aCuttingPositions[nCnt_Push].Y_Target THEN
					g_aCuttingPositions[nCnt_Push].bPushAwayProduct := FALSE;
					g_aCuttingPositions[nCnt_Push].rPushAwayDistance := 0;
				END_IF
			END_FOR
		END_IF
	END_IF

(**********************************************************************************************************************************
* Slab Triangle
**********************************************************************************************************************************)
ELSIF 	(g_HMI_RCP_Parameters.nProductType = Prod_Slab_Triangle_1x1) (*Horizontale component van nieuwe driehoeken*)
THEN

	rSizeOfKnife				:= g_HMI_MCH_Parameters.rSizeOfKnife;
	rCenterPointKnife			:= rSizeOfKnife/2;;
	rCenterPointKnifeInverted	:= rSizeOfKnife/2;;

	rProdLength_InY	:= g_HMI_RCP_Parameters.rProdLength_InY - MAX(0,g_HMI_RCP_Parameters.rSizeTrimRear) - MAX(0,g_HMI_RCP_Parameters.rSizeTrimFront);
	rProdLength_InX	:= g_HMI_RCP_Parameters.rProdLength_InX - MAX(0,g_HMI_RCP_Parameters.rSizeTrimRight) - MAX(0,g_HMI_RCP_Parameters.rSizeTrimLeft);

	(* Offset of slab *)
	FirstPoint.X	:= g_HMI_MCH_Parameters.rStartPointSlab_X;
	FirstPoint.Y	:= g_HMI_MCH_Parameters.rStartPointSlab_Y;

	rSizeTrimRear 	:= 	g_HMI_RCP_Parameters.rSizeTrimFront; (*AC 28-11-12: Omgedraaid vanaf HMI INstellingen*)
	rSizeTrimFront 	:= g_HMI_RCP_Parameters.rSizeTrimRear;(*AC 28-11-12: Omgedraaid vanaf HMI INstellingen*)
	rSizeTrimRight 	:= g_HMI_RCP_Parameters.rSizeTrimRight;
	rSizeTrimLeft 	:= g_HMI_RCP_Parameters.rSizeTrimLeft;

	(*g_rDistanceBetweenCuts_InY:=	(g_HMI_RCP_Parameters.rProdLength_InY - rSizeTrimRear - rSizeTrimFront) / INT_TO_REAL(g_HMI_RCP_Parameters.nPartsY);*)
	g_rDistanceBetweenCuts_InY	:= g_HMI_RCP_Parameters.rPartSizeY;
	g_sMACH.ERR.bPieceTooLarge := (rProdLength_InY < g_rDistanceBetweenCuts_InY) OR (rProdLength_InX < g_HMI_RCP_Parameters.rPartSizeX);

	(* Determine number of lines *)
	rNrOfLines	:=	(rProdLength_InY / g_rDistanceBetweenCuts_InY) - 1;
	nNrOfLines	:=	TRUNC_INT(rNrOfLines);
	IF	nNrOfLines < rNrOfLines	(* indien er nog product over is (afvalrand, dan aan weerszijden een afvalrand snijden *)
	THEN
		rWasteExtra := (rProdLength_InY - ((nNrOfLines +1)* g_rDistanceBetweenCuts_InY))/2;
		rSizeTrimRear	 	:= MAX(0,g_HMI_RCP_Parameters.rSizeTrimFront) + rWasteExtra;(*AC 28-11-12: Omgedraaid vanaf HMI INstellingen*)
		rSizeTrimFront 	:= MAX(0,g_HMI_RCP_Parameters.rSizeTrimRear) + rWasteExtra;
		g_bTrimRear		:= TRUE;
		g_bTrimFront		:= TRUE;
		nNrOfLines		:= nNrOfLines + 2;
	ELSE
		rSizeTrimRear	 	:= MAX(0, g_HMI_RCP_Parameters.rSizeTrimFront);(*AC 28-11-12: Omgedraaid vanaf HMI INstellingen*)
		rSizeTrimFront 	:= MAX(0, g_HMI_RCP_Parameters.rSizeTrimRear);(*AC 28-11-12: Omgedraaid vanaf HMI INstellingen*)
	END_IF
	(* Uitrekenen front en rear afvalrand *)
	rNrOfLines	:= (rProdLength_InX / g_rDistanceBetweenCuts_InX) - 1;
	nNrOfLines	:= TRUNC_INT(rNrOfLines);
	IF	nNrOfLines < rNrOfLines	(* indien er nog product over is (afvalrand, dan aan weerszijden een afvalrand snijden *)
	THEN
		rWasteExtra := (rProdLength_InX - ((nNrOfLines +1)* g_rDistanceBetweenCuts_InX))/2;
		rSizeTrimRight 	:= MAX(0,g_HMI_RCP_Parameters.rSizeTrimRight) + rWasteExtra;
		rSizeTrimLeft 	:= MAX(0,g_HMI_RCP_Parameters.rSizeTrimLeft) + rWasteExtra;
	ELSE
		rSizeTrimRight 	:= g_HMI_RCP_Parameters.rSizeTrimRight ;
		rSizeTrimLeft 	:= g_HMI_RCP_Parameters.rSizeTrimLeft;
	END_IF
	(* Determine number of lines *)
	rNrOfLines	:= (rProdLength_InY / g_rDistanceBetweenCuts_InY) - 1;
	nNrOfLines	:=	TRUNC_INT(rNrOfLines) + BOOL_TO_INT(rSizeTrimRear > 0) + BOOL_TO_INT(rSizeTrimFront > 0);

	overshootSettings.MarginXMin	:= C_rMinOvershootX;		(* Mechanical boundary *)
	overshootSettings.MarginXMax	:= SEL(gMachConfig.bXL,C_rMaxOvershootX,C_rMaxOvershootX_XL);	(* Mechanical boundary *)
	overshootSettings.MarginYMin	:= C_rMinOvershootY;		(* Mechanical boundary *)
	overshootSettings.MarginYMax	:= SEL(gMachConfig.bXL,C_rMaxOvershootY,C_rMaxOvershootY_XL);		(* Mechanical boundary *)

	overshootSettings.adjustXMax := TRUE;
	overshootSettings.adjustXMin := TRUE;
	overshootSettings.adjustYMax := TRUE;
	overshootSettings.adjustYMin := TRUE;

	(* Determine number of lines *)
	IF nNrOfLines > 0 THEN
		(* Calculate number of cuts on the line *)
		rLengthOfLine := g_HMI_RCP_Parameters.rProdLength_InX - rSizeTrimRight - rSizeTrimLeft;
		IF rLengthOfLine > rSizeOfKnife
		THEN
			nNumberOfCutsPerLine := TRUNC_INT(rLengthOfLine / rSizeOfKnife);
			IF nNumberOfCutsPerLine < (rLengthOfLine / rSizeOfKnife)
			THEN
				nNumberOfCutsPerLine := nNumberOfCutsPerLine + 1;
			END_IF
			rMmPerCut := (rLengthOfLine - rSizeOfKnife)/(nNumberOfCutsPerLine -1);
		ELSE
			nNumberOfCutsPerLine := 1;
		END_IF

		(* Calculate positions on first line *)
		IF g_bTrimRear
		THEN
			IF nNumberOfCutsPerLine = 1
			THEN
				IF NOT StorePos(I_rX:= 							FirstPoint.X + rSizeTrimRight + rCenterPointKnife,
								I_rY:=							(rFirstYPosition := FirstPoint.Y + rSizeTrimRear),
								I_rA:=							0,
								I_rK:=							0,
								I_bIsWaste :=					 (g_HMI_RCP_Parameters.bCutWasteFirst) ,
								I_sOvershootSettings := 		overshootSettings)
				THEN
										RETURN;
				END_IF

			ELSE
				FOR nCnt_pos:=1 TO (nNumberOfCutsPerLine - 1) DO
					IF NOT StorePos(I_rX:= 							FirstPoint.X + rSizeTrimRight + (nCnt_pos - 1) * rMmPerCut
																					 + rCenterPointKnife,
									I_rY:=							(rFirstYPosition := FirstPoint.Y + rSizeTrimRear),
									I_rA:=							0,
									I_rK:=							0,
									I_bIsWaste :=					 (g_HMI_RCP_Parameters.bCutWasteFirst) ,
									I_sOvershootSettings := 		overshootSettings)
					THEN
												RETURN;
					END_IF

				END_FOR
				(* Last position on the line *)
				IF NOT StorePos(I_rX:= 							FirstPoint.X + g_HMI_RCP_Parameters.rProdLength_InX - rSizeTrimLeft - rCenterPointKnifeInverted,
								I_rY:=							FirstPoint.Y + rSizeTrimRear,
								I_rA:=							0,
								I_rK:=							0,
								I_bIsWaste :=					 (g_HMI_RCP_Parameters.bCutWasteFirst) ,
								I_sOvershootSettings := 		overshootSettings)
				THEN
										RETURN;
				END_IF

			END_IF
		ELSE (* No waste strip at the left *)
			IF nNumberOfCutsPerLine = 1
			THEN
				IF NOT StorePos(I_rX:= 							FirstPoint.X + rSizeTrimRight + rCenterPointKnife,
								I_rY:=							(rFirstYPosition := FirstPoint.Y + rSizeTrimRear + g_rDistanceBetweenCuts_InY),
								I_rA:=							0,
								I_rK:=							0,
								I_bIsWaste :=					FALSE,
								I_sOvershootSettings := 		overshootSettings)
				THEN
										RETURN;
				END_IF

			ELSE
				FOR nCnt_pos:=1 TO (nNumberOfCutsPerLine - 1) DO
					IF NOT StorePos(I_rX:= 							FirstPoint.X + rSizeTrimRight + (nCnt_pos - 1) * rMmPerCut
																					 + rCenterPointKnife,
									I_rY:=							(rFirstYPosition := FirstPoint.Y + rSizeTrimRear + g_rDistanceBetweenCuts_InY),
									I_rA:=							0,
									I_rK:=							0,
									I_bIsWaste :=					FALSE,
									I_sOvershootSettings := 		overshootSettings)
					THEN
												RETURN;
					END_IF

				END_FOR
				(* Last position on the line *)
				IF NOT StorePos(I_rX:= 							FirstPoint.X + g_HMI_RCP_Parameters.rProdLength_InX - rSizeTrimLeft - rCenterPointKnifeInverted,
								I_rY:=							FirstPoint.Y + rSizeTrimRear + g_rDistanceBetweenCuts_InY,
								I_rA:=							0,
								I_rK:=							0,
								I_bIsWaste :=					FALSE,
								I_sOvershootSettings := 		overshootSettings)
				THEN
										RETURN;
				END_IF

			END_IF
		END_IF

		(* Fill in all other positions on the rest of the lines *)

		FOR nCnt_line := 2 TO (nNrOfLines) BY 1 DO
			IF nNumberOfCutsPerLine = 1
			THEN
				IF NOT StorePos(I_rX:= 							FirstPoint.X + rSizeTrimRight + rCenterPointKnife,
								I_rY:=							rFirstYPosition + (nCnt_line-1) * g_rDistanceBetweenCuts_InY,
								I_rA:=							0,
								I_rK:=							0,
								I_bIsWaste :=					 (g_HMI_RCP_Parameters.bCutWasteFirst AND g_bTrimFront AND nCnt_Line = nNrOfLines) ,
								I_sOvershootSettings := 		overshootSettings)
				THEN
										RETURN;
				END_IF

			ELSE
				IF bToggle (* from front to rear *)
				THEN
					FOR nCnt_pos:=1 TO (nNumberOfCutsPerLine - 1) DO
						IF NOT StorePos(I_rX:= 							FirstPoint.X + rSizeTrimRight + rCenterPointKnife
																                                                   + (nCnt_pos - 1) * rMmPerCut ,
										I_rY:=							rFirstYPosition + (nCnt_line-1) * g_rDistanceBetweenCuts_InY,
										I_rA:=							0,
										I_rK:=							0,
										I_bIsWaste :=					 (g_HMI_RCP_Parameters.bCutWasteFirst AND g_bTrimFront AND nCnt_Line = nNrOfLines) ,
										I_sOvershootSettings := 		overshootSettings)
						THEN
														RETURN;
						END_IF

					END_FOR
					(* Last position on the line *)
					IF NOT StorePos(I_rX:= 							FirstPoint.X + g_HMI_RCP_Parameters.rProdLength_InX - rSizeTrimLeft - rCenterPointKnifeInverted,
									I_rY:=							rFirstYPosition + (nCnt_line-1) * g_rDistanceBetweenCuts_InY,
									I_rA:=							0,
									I_rK:=							0,
									I_bIsWaste :=					 (g_HMI_RCP_Parameters.bCutWasteFirst AND g_bTrimFront AND nCnt_Line = nNrOfLines) ,
									I_sOvershootSettings := 		overshootSettings)
					THEN
												RETURN;
					END_IF

				ELSE (* toggle, ie from rear to front *)
					FOR nCnt_pos:=1 TO (nNumberOfCutsPerLine - 1) DO
						IF NOT StorePos(I_rX:= 							FirstPoint.X + g_HMI_RCP_Parameters.rProdLength_InX - rSizeTrimLeft - rCenterPointKnifeInverted
																							- (nCnt_pos -1) * rMmPerCut,
										I_rY:=							rFirstYPosition + (nCnt_line-1) * g_rDistanceBetweenCuts_InY,
										I_rA:=							0,
										I_rK:=							0,
										I_bIsWaste :=					 (g_HMI_RCP_Parameters.bCutWasteFirst AND g_bTrimFront AND nCnt_Line = nNrOfLines) ,
										I_sOvershootSettings := 		overshootSettings)
						THEN
														RETURN;
						END_IF

					END_FOR
					(* Last position on the line *)
					IF NOT StorePos(I_rX:= 							FirstPoint.X + rSizeTrimRight + rCenterPointKnife,
									I_rY:=							rFirstYPosition + (nCnt_line-1) * g_rDistanceBetweenCuts_InY,
									I_rA:=							0,
									I_rK:=							0,
									I_bIsWaste :=					 (g_HMI_RCP_Parameters.bCutWasteFirst AND g_bTrimFront AND nCnt_Line = nNrOfLines) ,
									I_sOvershootSettings := 		overshootSettings)
					THEN
												RETURN;
					END_IF

				END_IF
				bToggle := NOT bToggle;
			END_IF
		END_FOR

		(* Schuiven Uitbreiding AC *)
		(*Alle ingevulde posities controleren of Y gelijk is aan uiterste Y*)
		(*Indien ja: set bPushAwayProduct en corresponderende distance.*)
		IF g_bTrimFront THEN
			rLast_Y_Pos := rFirstYPosition + (nNrOfLines-1) * g_rDistanceBetweenCuts_InY;

			FOR nCnt_Push := nFirstPosFirstTray TO g_sCuttingPositionsInfo.index -1 DO
				IF rLast_Y_Pos = g_aCuttingPositions[nCnt_Push].Y_Target THEN
					g_aCuttingPositions[nCnt_Push].bPushAwayProduct := FALSE;
					g_aCuttingPositions[nCnt_Push].rPushAwayDistance := 0;
				END_IF
			END_FOR
		END_IF
	END_IF
(************************************************************************************************************
* Trays in triangle AC: 23-10-2012 -> EQUALS NORMAL SQUARE TRAY
****************************************************************************************************************)
END_IF

Calc_Hor := TRUE;

END_FUNCTION

(* ---- Calc_Round.fun ---- *)
FUNCTION Calc_Round : Bool
VAR_INPUT
	bIsLeftCake : BOOL;
	nPartsRound: INT;
	cutsToMake: INT;
	rSizeOfKnife				: REAL;
	rCutsPerLine				: REAL;
	rRotatiehoek: ARRAY[1..35] OF REAL;
	FirstPoint					: Gonio_Point;
	overshootSettings 			: Gonio_Settings;
END_VAR
VAR
	bToggle: BOOL;
	bKC1: BOOL;

	i: INT;
	c: INT;
	nCutsPerLine				: INT;

	rRotatiehoekInRad			: REAL;
	rDiameterTaart				: REAL;
	rKC2						: REAL;
	rStepDistX 					: REAL;
	rStepDistY 					: REAL;
END_VAR

	rDiameterTaart	:= g_HMI_RCP_Parameters.rDiameterRound;
	//nFirstPosFirstTray := g_sCuttingPositionsInfo.index;

	(*Calculate number of cuts*)
	rCutsPerLine := rDiameterTaart / rSizeOfKnife;
	nCutsPerLine := TRUNC_INT(rCutsPerLine);
	IF rCutsPerLine > nCutsPerLine THEN
		nCutsPerLine := nCutsPerLine + 1;
	END_IF

	IF bIsLeftCake THEN
		cutsToMake := Calc_RoundCakeDivisionsTable(I_Divisions:=g_HMI_RCP_Parameters.nPartsRound, I_InSequence := g_HMI_RCP_Parameters.bCutRoundInSequence, IQ_Table:= rRotatiehoek);
	ELSE
		cutsToMake := Calc_RoundCakeDivisionsTable(I_Divisions:=g_HMI_RCP_Parameters.nPartsRoundRight, I_InSequence := g_HMI_RCP_Parameters.bCutRoundInSequence, IQ_Table:= rRotatiehoek);
	END_IF

	IF (cutsToMake > 0) THEN

		FOR i :=1 TO (nPartsRound / 2) DO
			rRotatiehoekInRad	:=	(rRotatiehoek[i] / 360.0) * 2.0 * C_rPi;

			(*Verplaatsingen bepalen*)
			IF nCutsPerLine = 1 THEN
				rStepDistX := 0;
				rStepDistY := 0;
			ELSE
				rStepDistX := (rDiameterTaart - rSizeOfKnife)/(nCutsPerLine - 1)* COS(rRotatiehoekInRad);
				rStepDistY := (rDiameterTaart - rSizeOfKnife)/(nCutsPerLine - 1) * SIN(rRotatiehoekInRad);
			END_IF

			IF NOT bToggle THEN (* mes van MaxX/MinY naar MinX/MaxY*)
				FOR c := 0 TO nCutsPerLine-1 DO
					IF nCutsPerLine = 1 THEN
						IF NOT StorePos(I_rX:= 							FirstPoint.X + g_HMI_RCP_Parameters.rMidPosOffsetRound1X,
										I_rY:=							FirstPoint.Y + g_HMI_RCP_Parameters.rMidPosOffsetRound1Y,
										I_rA:=							rRotatiehoek[i],
										I_rK:=							0,
										I_bIsWaste :=					FALSE,
										I_sOvershootSettings := 		overshootSettings)
						THEN
										RETURN;
						END_IF
					ELSE
						IF NOT StorePos(I_rX:= 							FirstPoint.X + g_HMI_RCP_Parameters.rMidPosOffsetRound1X
																							+ (((rDiameterTaart - rSizeOfKnife) / 2) * COS(rRotatiehoekInRad))
																							- (c * rStepDistX),
										I_rY:=							FirstPoint.Y + g_HMI_RCP_Parameters.rMidPosOffsetRound1Y
																							+ (((rDiameterTaart - rSizeOfKnife) / 2) * SIN(rRotatiehoekInRad))
																							- (c * rStepDistY),
										I_rA:=							rRotatiehoek[i],
										I_rK:=							0,
										I_bIsWaste :=					FALSE,
										I_sOvershootSettings := 		overshootSettings)
						THEN
										RETURN;
						END_IF
					END_IF
				END_FOR
			ELSE (* toggle, mes van linksonder naar rechtsboven *)
				FOR c := 0 TO nCutsPerLine-1 DO
					IF nCutsPerLine = 1 THEN
						IF NOT StorePos(I_rX:= 							FirstPoint.X + g_HMI_RCP_Parameters.rMidPosOffsetRound1X,
										I_rY:=							FirstPoint.Y + g_HMI_RCP_Parameters.rMidPosOffsetRound1Y,
										I_rA:=							rRotatiehoek[i],
										I_rK:=							0,
										I_bIsWaste :=					FALSE,
										I_sOvershootSettings := 		overshootSettings)
						THEN
										RETURN;
						END_IF

					ELSE
						IF NOT StorePos(I_rX:= 							FirstPoint.X + g_HMI_RCP_Parameters.rMidPosOffsetRound1X
																								- (((rDiameterTaart - rSizeOfKnife) / 2) * COS(rRotatiehoekInRad))
																								+ (c * rStepDistX),
										I_rY:=							FirstPoint.Y + g_HMI_RCP_Parameters.rMidPosOffsetRound1Y
																								- (((rDiameterTaart - rSizeOfKnife) / 2) * SIN(rRotatiehoekInRad))
																								+ (c * rStepDistY),
										I_rA:=							rRotatiehoek[i],
										I_rK:=							0,
										I_bIsWaste :=					FALSE,
										I_sOvershootSettings := 		overshootSettings)
						THEN
										RETURN;
						END_IF
						IF g_sCuttingPositionsInfo.index = 4 THEN bKC1 := TRUE; rKC2 := COS(90); END_IF
					END_IF
				END_FOR
			END_IF
			bToggle := NOT bToggle;
		END_FOR
	END_IF

END_FUNCTION

(* ---- Calc_RoundCakeDivisionsTable.fun ---- *)
FUNCTION Calc_RoundCakeDivisionsTable : INT
VAR_INPUT
	I_Divisions		: INT;
	I_InSequence	: BOOL;
END_VAR
VAR_IN_OUT
	IQ_Table		: ARRAY[*] OF REAL;
END_VAR
VAR
	i				: INT;
	lower			: DINT;
	upper 			: DINT;
END_VAR

(*
	Fills the array IQ_Table table with the rotations in degrees in order to cut in I_Divisions pieces.
	Returns an integer representing how many cuts to place.
	Returns -1 if an error occured.
*)

lower := LOWER_BOUND(IQ_Table,1);
upper := UPPER_BOUND(IQ_Table,1);

IF (I_Divisions > 70 OR I_Divisions < 2) THEN
	//Hardcoded limit to make sure we dont cut the cake to pulp or dont cut at all.
	Calc_RoundCakeDivisionsTable := -1;
	RETURN;
END_IF

IF (I_Divisions MOD 2) > 0 THEN
	//Uneven number of cuts.
	Calc_RoundCakeDivisionsTable := -1;
	RETURN;
END_IF

IF (I_Divisions / 2) > (upper - lower) THEN
	//We cant store this many cuts in the table.
	Calc_RoundCakeDivisionsTable := -1;
	RETURN;
END_IF

IF I_InSequence THEN
	FOR i := 0 TO (I_Divisions/2) DO
		IQ_Table[i + lower] := i * (360.0/INT_TO_REAL(I_Divisions));
	END_FOR
ELSE

	CASE I_Divisions OF
		2:
			IQ_Table[ lower + 0] := 0;

		4:
			IQ_Table[ lower + 0] := 0;
			IQ_Table[ lower + 1] := 90;

		6:
			IQ_Table[ lower + 0] := 0;
			IQ_Table[ lower + 1] := 60;
			IQ_Table[ lower + 2] := 120;

		8:
			IQ_Table[ lower + 0] := 0;
			IQ_Table[ lower + 1] := 90;
			IQ_Table[ lower + 2] := 45;
			IQ_Table[ lower + 3] := 135;

		10:
			IQ_Table[ lower + 0] := 0;
			IQ_Table[ lower + 1] := 108;
			IQ_Table[ lower + 2] := 36;
			IQ_Table[ lower + 3] := 144;
			IQ_Table[ lower + 4] := 72;

		12:
			IQ_Table[ lower + 0] := 0;
			IQ_Table[ lower + 1] := 90;
			IQ_Table[ lower + 2] := 120;
			IQ_Table[ lower + 3] := 60;
			IQ_Table[ lower + 4] := 30;
			IQ_Table[ lower + 5] := 150;

		14:
			IQ_Table[ lower + 0] := 0;
			IQ_Table[ lower + 1] := 102.86;
			IQ_Table[ lower + 2] := 51.43;
			IQ_Table[ lower + 3] := 128.57;
			IQ_Table[ lower + 4] := 77.14;
			IQ_Table[ lower + 5] := 25.71;
			IQ_Table[ lower + 6] := 154.29;

		(* Nieuw voor Smaak & Co *)
		16:
			IQ_Table[ lower + 0] := 0;
			IQ_Table[ lower + 1] := 90;
			IQ_Table[ lower + 2] := 45;
			IQ_Table[ lower + 3] := 135;
			IQ_Table[ lower + 4] := 22.5;
			IQ_Table[ lower + 5] := 112.5;
			IQ_Table[ lower + 6] := 67.5;
			IQ_Table[ lower + 7] := 157.5;

		18:
			IQ_Table[ lower + 0] := 0;
			IQ_Table[ lower + 1] := 80;
			IQ_Table[ lower + 2] := 40;
			IQ_Table[ lower + 3] := 120;
			IQ_Table[ lower + 4] := 20;
			IQ_Table[ lower + 5] := 100;
			IQ_Table[ lower + 6] := 60;
			IQ_Table[ lower + 7] := 160;
			IQ_Table[ lower + 8] := 140;

		20:
			IQ_Table[ lower + 0] := 0;
			IQ_Table[ lower + 1] := 90;
			IQ_Table[ lower + 2] := 36;
			IQ_Table[ lower + 3] := 126;
			IQ_Table[ lower + 4] := 72;
			IQ_Table[ lower + 5] := 144;
			IQ_Table[ lower + 6] := 54;
			IQ_Table[ lower + 7] := 162;
			IQ_Table[ lower + 8] := 18;
			IQ_Table[ lower + 9] := 108;

		22:
			IQ_Table[ lower + 0] := 0;
			IQ_Table[ lower + 1] := 81.82;
			IQ_Table[ lower + 2] := 130.91;
			IQ_Table[ lower + 3] := 49.09;
			IQ_Table[ lower + 4] := 147.27;
			IQ_Table[ lower + 5] := 65.45;
			IQ_Table[ lower + 6] := 32.73;
			IQ_Table[ lower + 7] := 98.18;
			IQ_Table[ lower + 8] := 163.64;
			IQ_Table[ lower + 9] := 114.55;
			IQ_Table[ lower + 10] := 16.36;

		24:
			IQ_Table[ lower + 0] := 0;
			IQ_Table[ lower + 1] := 90;
			IQ_Table[ lower + 2] := 45;
			IQ_Table[ lower + 3] := 135;
			IQ_Table[ lower + 4] := 165;
			IQ_Table[ lower + 5] := 75;
			IQ_Table[ lower + 6] := 120;
			IQ_Table[ lower + 7] := 30;
			IQ_Table[ lower + 8] := 60;
			IQ_Table[ lower + 9] := 150;
			IQ_Table[ lower + 10] := 105;
			IQ_Table[ lower + 11] := 15;

		26:
			IQ_Table[ lower + 0] := 0;
			IQ_Table[ lower + 1] := 96.92;
			IQ_Table[ lower + 2] := 41.54;
			IQ_Table[ lower + 3] := 138.46;
			IQ_Table[ lower + 4] := 69.23;
			IQ_Table[ lower + 5] := 166.15;
			IQ_Table[ lower + 6] := 27.69;
			IQ_Table[ lower + 7] := 110.77;
			IQ_Table[ lower + 8] := 55.38;
			IQ_Table[ lower + 9] := 124.62;
			IQ_Table[ lower + 10] := 83.08;
			IQ_Table[ lower + 11] := 152.31;
			IQ_Table[ lower + 12] := 13.85;

		28:
			IQ_Table[ lower + 0] := 0;
			IQ_Table[ lower + 1] := 90;
			IQ_Table[ lower + 2] := 128.57;
			IQ_Table[ lower + 3] := 38.57;
			IQ_Table[ lower + 4] := 167.14;
			IQ_Table[ lower + 5] := 64.29;
			IQ_Table[ lower + 6] := 25.71;
			IQ_Table[ lower + 7] := 141.43;
			IQ_Table[ lower + 8] := 102.86;
			IQ_Table[ lower + 9] := 77.14;
			IQ_Table[ lower + 10] := 154.29;
			IQ_Table[ lower + 11] := 51.43;
			IQ_Table[ lower + 12] := 115.71;
			IQ_Table[ lower + 13] := 12.86;

		30:
			IQ_Table[ lower + 0] := 0.00;
			IQ_Table[ lower + 1] := 84.00;
			IQ_Table[ lower + 2] := 48.00;
			IQ_Table[ lower + 3] := 132.00;
			IQ_Table[ lower + 4] := 24.00;
			IQ_Table[ lower + 5] := 108.00;
			IQ_Table[ lower + 6] := 60.00;
			IQ_Table[ lower + 7] := 144.00;
			IQ_Table[ lower + 8] := 12.00;
			IQ_Table[ lower + 9] := 72.00;
			IQ_Table[ lower + 10] := 120.00;
			IQ_Table[ lower + 11] := 36.00;
			IQ_Table[ lower + 12] := 156.00;
			IQ_Table[ lower + 13] := 96.00;
			IQ_Table[ lower + 14] := 168.00;

		32:
			IQ_Table[ lower + 0] := 0.00;
			IQ_Table[ lower + 1] := 90.00;
			IQ_Table[ lower + 2] := 45.00;
			IQ_Table[ lower + 3] := 135.00;
			IQ_Table[ lower + 4] := 22.50;
			IQ_Table[ lower + 5] := 67.50;
			IQ_Table[ lower + 6] := 112.50;
			IQ_Table[ lower + 7] := 157.50;
			IQ_Table[ lower + 8] := 33.75;
			IQ_Table[ lower + 9] := 78.75;
			IQ_Table[ lower + 10] := 123.75;
			IQ_Table[ lower + 11] := 168.75;
			IQ_Table[ lower + 12] := 11.25;
			IQ_Table[ lower + 13] := 56.25;
			IQ_Table[ lower + 14] := 101.25;
			IQ_Table[ lower + 15] := 146.25;

		34:
			IQ_Table[ lower + 0] := 0.00;
			IQ_Table[ lower + 1] := 84.71;
			IQ_Table[ lower + 2] := 42.35;
			IQ_Table[ lower + 3] := 137.65;
			IQ_Table[ lower + 4] := 21.18;
			IQ_Table[ lower + 5] := 63.53;
			IQ_Table[ lower + 6] := 116.47;
			IQ_Table[ lower + 7] := 158.82;
			IQ_Table[ lower + 8] := 31.76;
			IQ_Table[ lower + 9] := 105.88;
			IQ_Table[ lower + 10] := 74.12;
			IQ_Table[ lower + 11] := 148.24;
			IQ_Table[ lower + 12] := 10.59;
			IQ_Table[ lower + 13] := 52.94;
			IQ_Table[ lower + 14] := 95.29;
			IQ_Table[ lower + 15] := 127.06;
			IQ_Table[ lower + 16] := 169.41;

		36:
			IQ_Table[ lower + 0] := 0.00;
			IQ_Table[ lower + 1] := 90.00;
			IQ_Table[ lower + 2] := 40.00;
			IQ_Table[ lower + 3] := 130.00;
			IQ_Table[ lower + 4] := 20.00;
			IQ_Table[ lower + 5] := 110.00;
			IQ_Table[ lower + 6] := 60.00;
			IQ_Table[ lower + 7] := 150.00;
			IQ_Table[ lower + 8] := 30.00;
			IQ_Table[ lower + 9] := 120.00;
			IQ_Table[ lower + 10] := 70.00;
			IQ_Table[ lower + 11] := 160.00;
			IQ_Table[ lower + 12] := 10.00;
			IQ_Table[ lower + 13] := 100.00;
			IQ_Table[ lower + 14] := 50.00;
			IQ_Table[ lower + 15] := 140.00;
			IQ_Table[ lower + 16] := 80.00;
			IQ_Table[ lower + 17] := 170.00;

		38:
			IQ_Table[ lower + 0] := 0.00;
			IQ_Table[ lower + 1] := 85.26;
			IQ_Table[ lower + 2] := 47.37;
			IQ_Table[ lower + 3] := 132.63;
			IQ_Table[ lower + 4] := 28.42;
			IQ_Table[ lower + 5] := 113.68;
			IQ_Table[ lower + 6] := 66.32;
			IQ_Table[ lower + 7] := 161.05;
			IQ_Table[ lower + 8] := 9.47;
			IQ_Table[ lower + 9] := 104.21;
			IQ_Table[ lower + 10] := 56.84;
			IQ_Table[ lower + 11] := 142.11;
			IQ_Table[ lower + 12] := 75.79;
			IQ_Table[ lower + 13] := 170.53;
			IQ_Table[ lower + 14] := 18.95;
			IQ_Table[ lower + 15] := 123.16;
			IQ_Table[ lower + 16] := 37.89;
			IQ_Table[ lower + 17] := 94.74;
			IQ_Table[ lower + 18] := 151.58;

		40:
			IQ_Table[ lower + 0]  := 0;
			IQ_Table[ lower + 1]  := 90.00;
			IQ_Table[ lower + 2]  := 45.00;
			IQ_Table[ lower + 3]  := 135.00;
			IQ_Table[ lower + 4]  := 27.00;
			IQ_Table[ lower + 5]  := 117.00;
			IQ_Table[ lower + 6]  := 72.00;
			IQ_Table[ lower + 7]  := 162.00;
			IQ_Table[ lower + 8]  := 36.00;
			IQ_Table[ lower + 9] := 126.00;
			IQ_Table[ lower + 10] := 63.00;
			IQ_Table[ lower + 11] := 153.00;
			IQ_Table[ lower + 12] := 18.00;
			IQ_Table[ lower + 13] := 108.00;
			IQ_Table[ lower + 14] := 54.00;
			IQ_Table[ lower + 15] := 144.00;
			IQ_Table[ lower + 16] := 9.00;
			IQ_Table[ lower + 17] := 99.00;
			IQ_Table[ lower + 18] := 81.00;
			IQ_Table[ lower + 19] := 171.00;

		42:
			IQ_Table[ lower + 0]  := 0;
			IQ_Table[ lower + 1]  := 85.71;
			IQ_Table[ lower + 2]  := 42.86;
			IQ_Table[ lower + 3]  := 137.14;
			IQ_Table[ lower + 4]  := 25.71;
			IQ_Table[ lower + 5]  := 111.43;
			IQ_Table[ lower + 6]  := 68.57;
			IQ_Table[ lower + 7]  := 162.86;
			IQ_Table[ lower + 8]  := 17.14;
			IQ_Table[ lower + 9] := 102.86;
			IQ_Table[ lower + 10] := 51.43;
			IQ_Table[ lower + 11] := 145.71;
			IQ_Table[ lower + 12] := 34.29;
			IQ_Table[ lower + 13] := 120.00;
			IQ_Table[ lower + 14] := 60.00;
			IQ_Table[ lower + 15] := 154.29;
			IQ_Table[ lower + 16] := 77.14;
			IQ_Table[ lower + 17] := 128.57;
			IQ_Table[ lower + 18] := 8.57;
			IQ_Table[ lower + 19] := 94.29;
			IQ_Table[ lower + 20] := 171.43;

		44:
			IQ_Table[ lower + 0]  := 0;
			IQ_Table[ lower + 1]  := 90.00;
			IQ_Table[ lower + 2]  := 40.91;
			IQ_Table[ lower + 3]  := 130.91;
			IQ_Table[ lower + 4]  := 65.45;
			IQ_Table[ lower + 5]  := 155.45;
			IQ_Table[ lower + 6]  := 24.55;
			IQ_Table[ lower + 7]  := 114.55;
			IQ_Table[ lower + 8]  := 49.09;
			IQ_Table[ lower + 9] := 139.09;
			IQ_Table[ lower + 10] := 16.36;
			IQ_Table[ lower + 11] := 106.36;
			IQ_Table[ lower + 12] := 57.27;
			IQ_Table[ lower + 13] := 147.27;
			IQ_Table[ lower + 14] := 8.18;
			IQ_Table[ lower + 15] := 98.18;
			IQ_Table[ lower + 16] := 73.64;
			IQ_Table[ lower + 17] := 163.64;
			IQ_Table[ lower + 18] := 32.73;
			IQ_Table[ lower + 19] := 122.73;
			IQ_Table[ lower + 20] := 81.82;
			IQ_Table[ lower + 21] := 171.82;

		46:
			IQ_Table[ lower + 0]  := 0;
			IQ_Table[ lower + 1]  := 93.91;
			IQ_Table[ lower + 2]  := 46.96;
			IQ_Table[ lower + 3]  := 133.04;
			IQ_Table[ lower + 4]  := 23.48;
			IQ_Table[ lower + 5]  := 117.39;
			IQ_Table[ lower + 6]  := 70.43;
			IQ_Table[ lower + 7]  := 156.52;
			IQ_Table[ lower + 8]  := 31.30;
			IQ_Table[ lower + 9] := 125.22;
			IQ_Table[ lower + 10] := 62.61;
			IQ_Table[ lower + 11] := 148.70;
			IQ_Table[ lower + 12] := 15.65;
			IQ_Table[ lower + 13] := 109.57;
			IQ_Table[ lower + 14] := 54.78;
			IQ_Table[ lower + 15] := 140.87;
			IQ_Table[ lower + 16] := 86.09;
			IQ_Table[ lower + 17] := 172.17;
			IQ_Table[ lower + 18] := 39.13;
			IQ_Table[ lower + 19] := 101.74;
			IQ_Table[ lower + 20] := 7.83;
			IQ_Table[ lower + 21] := 78.26;
			IQ_Table[ lower + 22] := 164.35;

		48:
			IQ_Table[ lower + 0]  := 0;
			IQ_Table[ lower + 1]  := 90.00;
			IQ_Table[ lower + 2]  := 45.00;
			IQ_Table[ lower + 3]  := 135.00;
			IQ_Table[ lower + 4]  := 22.50;
			IQ_Table[ lower + 5]  := 112.50;
			IQ_Table[ lower + 6]  := 67.50;
			IQ_Table[ lower + 7]  := 157.50;
			IQ_Table[ lower + 8]  := 15.00;
			IQ_Table[ lower + 9] := 105.00;
			IQ_Table[ lower + 10] := 52.50;
			IQ_Table[ lower + 11] := 142.50;
			IQ_Table[ lower + 12] := 30.00;
			IQ_Table[ lower + 13] := 120.00;
			IQ_Table[ lower + 14] := 82.50;
			IQ_Table[ lower + 15] := 172.50;
			IQ_Table[ lower + 16] := 37.50;
			IQ_Table[ lower + 17] := 127.50;
			IQ_Table[ lower + 18] := 60.00;
			IQ_Table[ lower + 19] := 150.00;
			IQ_Table[ lower + 20] := 7.50;
			IQ_Table[ lower + 21] := 97.50;
			IQ_Table[ lower + 22] := 75.00;
			IQ_Table[ lower + 23] := 165.00;

		50:
			IQ_Table[ lower + 0]  := 0.00;
			IQ_Table[ lower + 1]  := 93.60;
			IQ_Table[ lower + 2]  := 43.20;
			IQ_Table[ lower + 3]  := 136.80;
			IQ_Table[ lower + 4]  := 21.60;
			IQ_Table[ lower + 5]  := 72.00;
			IQ_Table[ lower + 6]  := 115.20;
			IQ_Table[ lower + 7]  := 158.40;
			IQ_Table[ lower + 8]  := 7.20;
			IQ_Table[ lower + 9]  := 100.80;
			IQ_Table[ lower + 10]  := 57.60;
			IQ_Table[ lower + 11]  := 151.20;
			IQ_Table[ lower + 12]  := 36.00;
			IQ_Table[ lower + 13]  := 122.40;
			IQ_Table[ lower + 14]  := 64.80;
			IQ_Table[ lower + 15]  := 165.60;
			IQ_Table[ lower + 16]  := 14.40;
			IQ_Table[ lower + 17]  := 86.40;
			IQ_Table[ lower + 18]  := 50.40;
			IQ_Table[ lower + 19]  := 144.00;
			IQ_Table[ lower + 20]  := 79.20;
			IQ_Table[ lower + 21]  := 108.00;
			IQ_Table[ lower + 22]  := 172.80;
			IQ_Table[ lower + 23]  := 28.80;
			IQ_Table[ lower + 24]  := 129.60;

		52:
			IQ_Table[ lower + 0]  := 0.00;
			IQ_Table[ lower + 1]  := 90.00;
			IQ_Table[ lower + 2]  := 48.46;
			IQ_Table[ lower + 3]  := 138.46;
			IQ_Table[ lower + 4]  := 27.69;
			IQ_Table[ lower + 5]  := 117.69;
			IQ_Table[ lower + 6]  := 69.23;
			IQ_Table[ lower + 7]  := 159.23;
			IQ_Table[ lower + 8]  := 13.85;
			IQ_Table[ lower + 9]  := 103.85;
			IQ_Table[ lower + 10]  := 55.38;
			IQ_Table[ lower + 11]  := 145.38;
			IQ_Table[ lower + 12]  := 20.77;
			IQ_Table[ lower + 13]  := 110.77;
			IQ_Table[ lower + 14]  := 76.15;
			IQ_Table[ lower + 15]  := 166.15;
			IQ_Table[ lower + 16]  := 6.92;
			IQ_Table[ lower + 17]  := 96.92;
			IQ_Table[ lower + 18]  := 41.54;
			IQ_Table[ lower + 19]  := 131.54;
			IQ_Table[ lower + 20]  := 62.31;
			IQ_Table[ lower + 21]  := 152.31;
			IQ_Table[ lower + 22]  := 34.62;
			IQ_Table[ lower + 23]  := 124.62;
			IQ_Table[ lower + 24]  := 83.08;
			IQ_Table[ lower + 25]  := 173.08;

		54:
			IQ_Table[ lower + 0]  := 0.00;
			IQ_Table[ lower + 1]  := 86.67;
			IQ_Table[ lower + 2]  := 46.67;
			IQ_Table[ lower + 3]  := 133.33;
			IQ_Table[ lower + 4]  := 26.67;
			IQ_Table[ lower + 5]  := 113.33;
			IQ_Table[ lower + 6]  := 66.67;
			IQ_Table[ lower + 7]  := 153.33;
			IQ_Table[ lower + 8]  := 13.33;
			IQ_Table[ lower + 9]  := 100.00;
			IQ_Table[ lower + 10]  := 53.33;
			IQ_Table[ lower + 11]  := 146.67;
			IQ_Table[ lower + 12]  := 33.33;
			IQ_Table[ lower + 13]  := 120.00;
			IQ_Table[ lower + 14]  := 60.00;
			IQ_Table[ lower + 15]  := 160.00;
			IQ_Table[ lower + 16]  := 6.67;
			IQ_Table[ lower + 17]  := 93.33;
			IQ_Table[ lower + 18]  := 40.00;
			IQ_Table[ lower + 19]  := 140.00;
			IQ_Table[ lower + 20]  := 20.00;
			IQ_Table[ lower + 21]  := 80.00;
			IQ_Table[ lower + 22]  := 166.67;
			IQ_Table[ lower + 23]  := 73.33;
			IQ_Table[ lower + 24]  := 106.67;
			IQ_Table[ lower + 25]  := 173.33;
			IQ_Table[ lower + 26]  := 126.67;

		56:
			IQ_Table[ lower + 0]  := 0.00;
			IQ_Table[ lower + 1]  := 90.00;
			IQ_Table[ lower + 2]  := 45.00;
			IQ_Table[ lower + 3]  := 135.00;
			IQ_Table[ lower + 4]  := 25.71;
			IQ_Table[ lower + 5]  := 115.71;
			IQ_Table[ lower + 6]  := 70.71;
			IQ_Table[ lower + 7]  := 160.71;
			IQ_Table[ lower + 8]  := 12.86;
			IQ_Table[ lower + 9]  := 102.86;
			IQ_Table[ lower + 10]  := 57.86;
			IQ_Table[ lower + 11]  := 147.86;
			IQ_Table[ lower + 12]  := 38.57;
			IQ_Table[ lower + 13]  := 128.57;
			IQ_Table[ lower + 14]  := 83.57;
			IQ_Table[ lower + 15]  := 173.57;
			IQ_Table[ lower + 16]  := 6.43;
			IQ_Table[ lower + 17]  := 96.43;
			IQ_Table[ lower + 18]  := 51.43;
			IQ_Table[ lower + 19]  := 141.43;
			IQ_Table[ lower + 20]  := 32.14;
			IQ_Table[ lower + 21]  := 122.14;
			IQ_Table[ lower + 22]  := 64.29;
			IQ_Table[ lower + 23]  := 154.29;
			IQ_Table[ lower + 24]  := 19.29;
			IQ_Table[ lower + 25]  := 109.29;
			IQ_Table[ lower + 26]  := 77.14;
			IQ_Table[ lower + 27]  := 167.14;

		58:
			IQ_Table[ lower + 0]  := 0.00;
			IQ_Table[ lower + 1]  := 93.10;
			IQ_Table[ lower + 2]  := 43.45;
			IQ_Table[ lower + 3]  := 136.55;
			IQ_Table[ lower + 4]  := 24.83;
			IQ_Table[ lower + 5]  := 117.93;
			IQ_Table[ lower + 6]  := 68.28;
			IQ_Table[ lower + 7]  := 161.38;
			IQ_Table[ lower + 8]  := 37.24;
			IQ_Table[ lower + 9]  := 130.34;
			IQ_Table[ lower + 10]  := 55.86;
			IQ_Table[ lower + 11]  := 148.97;
			IQ_Table[ lower + 12]  := 12.41;
			IQ_Table[ lower + 13]  := 105.52;
			IQ_Table[ lower + 14]  := 31.03;
			IQ_Table[ lower + 15]  := 124.14;
			IQ_Table[ lower + 16]  := 49.66;
			IQ_Table[ lower + 17]  := 142.76;
			IQ_Table[ lower + 18]  := 6.21;
			IQ_Table[ lower + 19]  := 99.31;
			IQ_Table[ lower + 20]  := 62.07;
			IQ_Table[ lower + 21]  := 155.17;
			IQ_Table[ lower + 22]  := 74.48;
			IQ_Table[ lower + 23]  := 111.72;
			IQ_Table[ lower + 24]  := 173.79;
			IQ_Table[ lower + 25]  := 86.90;
			IQ_Table[ lower + 26]  := 18.62;
			IQ_Table[ lower + 27]  := 167.59;
			IQ_Table[ lower + 28]  := 80.69;

		60:
			IQ_Table[ lower + 0]  := 0.00;
			IQ_Table[ lower + 1]  := 90.00;
			IQ_Table[ lower + 2]  := 48.00;
			IQ_Table[ lower + 3]  := 138.00;
			IQ_Table[ lower + 4]  := 24.00;
			IQ_Table[ lower + 5]  := 114.00;
			IQ_Table[ lower + 6]  := 66.00;
			IQ_Table[ lower + 7]  := 156.00;
			IQ_Table[ lower + 8]  := 36.00;
			IQ_Table[ lower + 9]  := 126.00;
			IQ_Table[ lower + 10]  := 78.00;
			IQ_Table[ lower + 11]  := 168.00;
			IQ_Table[ lower + 12]  := 12.00;
			IQ_Table[ lower + 13]  := 102.00;
			IQ_Table[ lower + 14]  := 60.00;
			IQ_Table[ lower + 15]  := 150.00;
			IQ_Table[ lower + 16]  := 30.00;
			IQ_Table[ lower + 17]  := 120.00;
			IQ_Table[ lower + 18]  := 72.00;
			IQ_Table[ lower + 19]  := 162.00;
			IQ_Table[ lower + 20]  := 6.00;
			IQ_Table[ lower + 21]  := 96.00;
			IQ_Table[ lower + 22]  := 42.00;
			IQ_Table[ lower + 23]  := 132.00;
			IQ_Table[ lower + 24]  := 18.00;
			IQ_Table[ lower + 25]  := 108.00;
			IQ_Table[ lower + 26]  := 54.00;
			IQ_Table[ lower + 27]  := 144.00;
			IQ_Table[ lower + 28]  := 84.00;
			IQ_Table[ lower + 29]  := 174.00;

		62:
			IQ_Table[ lower + 0]  := 0.00;
			IQ_Table[ lower + 1]  := 92.90;
			IQ_Table[ lower + 2]  := 46.45;
			IQ_Table[ lower + 3]  := 139.35;
			IQ_Table[ lower + 4]  := 29.03;
			IQ_Table[ lower + 5]  := 116.13;
			IQ_Table[ lower + 6]  := 69.68;
			IQ_Table[ lower + 7]  := 156.77;
			IQ_Table[ lower + 8]  := 11.61;
			IQ_Table[ lower + 9]  := 104.52;
			IQ_Table[ lower + 10]  := 52.26;
			IQ_Table[ lower + 11]  := 145.16;
			IQ_Table[ lower + 12]  := 23.23;
			IQ_Table[ lower + 13]  := 110.32;
			IQ_Table[ lower + 14]  := 40.65;
			IQ_Table[ lower + 15]  := 133.55;
			IQ_Table[ lower + 16]  := 5.81;
			IQ_Table[ lower + 17]  := 87.10;
			IQ_Table[ lower + 18]  := 58.06;
			IQ_Table[ lower + 19]  := 162.58;
			IQ_Table[ lower + 20]  := 34.84;
			IQ_Table[ lower + 21]  := 127.74;
			IQ_Table[ lower + 22]  := 75.48;
			IQ_Table[ lower + 23]  := 168.39;
			IQ_Table[ lower + 24]  := 17.42;
			IQ_Table[ lower + 25]  := 98.71;
			IQ_Table[ lower + 26]  := 63.87;
			IQ_Table[ lower + 27]  := 150.97;
			IQ_Table[ lower + 28]  := 121.94;
			IQ_Table[ lower + 29]  := 174.19;
			IQ_Table[ lower + 30]  := 81.29;

		64:
			IQ_Table[ lower + 0]  := 0;
			IQ_Table[ lower + 1]  := 90;
			IQ_Table[ lower + 2]  := 45;
			IQ_Table[ lower + 3]  := 135;
			IQ_Table[ lower + 4]  := 22.5;
			IQ_Table[ lower + 5]  := 112.5;
			IQ_Table[ lower + 6]  := 67.5;
			IQ_Table[ lower + 7]  := 157.5;
			IQ_Table[ lower + 8]  := 11.25;
			IQ_Table[ lower + 9]  := 101.25;
			IQ_Table[ lower + 10]  := 56.25;
			IQ_Table[ lower + 11]  := 146.25;
			IQ_Table[ lower + 12]  := 78.75;
			IQ_Table[ lower + 13]  := 168.75;
			IQ_Table[ lower + 14]  := 33.75;
			IQ_Table[ lower + 15]  := 123.75;
			IQ_Table[ lower + 16]  := 61.875;
			IQ_Table[ lower + 17]  := 151.875;
			IQ_Table[ lower + 18]  := 28.125;
			IQ_Table[ lower + 19]  := 118.125;
			IQ_Table[ lower + 20]  := 50.625;
			IQ_Table[ lower + 21]  := 140.625;
			IQ_Table[ lower + 22]  := 5.625;
			IQ_Table[ lower + 23]  := 95.625;
			IQ_Table[ lower + 24]  := 39.375;
			IQ_Table[ lower + 25]  := 129.375;
			IQ_Table[ lower + 26]  := 16.875;
			IQ_Table[ lower + 27]  := 106.875;
			IQ_Table[ lower + 28]  := 73.125;
			IQ_Table[ lower + 29]  := 163.125;
			IQ_Table[ lower + 30]  := 84.375;
			IQ_Table[ lower + 31]  := 174.375;

		66:
			IQ_Table[ lower + 0]  := 0.00;
			IQ_Table[ lower + 1]  := 87.27;
			IQ_Table[ lower + 2]  := 43.64;
			IQ_Table[ lower + 3]  := 136.36;
			IQ_Table[ lower + 4]  := 16.36;
			IQ_Table[ lower + 5]  := 109.09;
			IQ_Table[ lower + 6]  := 65.45;
			IQ_Table[ lower + 7]  := 158.18;
			IQ_Table[ lower + 8]  := 32.73;
			IQ_Table[ lower + 9]  := 125.45;
			IQ_Table[ lower + 10]  := 76.36;
			IQ_Table[ lower + 11]  := 169.09;
			IQ_Table[ lower + 12]  := 21.82;
			IQ_Table[ lower + 13]  := 114.55;
			IQ_Table[ lower + 14]  := 54.55;
			IQ_Table[ lower + 15]  := 147.27;
			IQ_Table[ lower + 16]  := 5.45;
			IQ_Table[ lower + 17]  := 98.18;
			IQ_Table[ lower + 18]  := 49.09;
			IQ_Table[ lower + 19]  := 141.82;
			IQ_Table[ lower + 20]  := 27.27;
			IQ_Table[ lower + 21]  := 120.00;
			IQ_Table[ lower + 22]  := 70.91;
			IQ_Table[ lower + 23]  := 163.64;
			IQ_Table[ lower + 24]  := 10.91;
			IQ_Table[ lower + 25]  := 103.64;
			IQ_Table[ lower + 26]  := 60.00;
			IQ_Table[ lower + 27]  := 152.73;
			IQ_Table[ lower + 28]  := 174.55;
			IQ_Table[ lower + 29]  := 92.73;
			IQ_Table[ lower + 30]  := 130.91;
			IQ_Table[ lower + 31]  := 81.82;
			IQ_Table[ lower + 32]  := 38.18;

		68:
			IQ_Table[ lower + 0]  := 0.00;
			IQ_Table[ lower + 1]  := 90.00;
			IQ_Table[ lower + 2]  := 47.65;
			IQ_Table[ lower + 3]  := 137.65;
			IQ_Table[ lower + 4]  := 21.18;
			IQ_Table[ lower + 5]  := 116.47;
			IQ_Table[ lower + 6]  := 68.82;
			IQ_Table[ lower + 7]  := 158.82;
			IQ_Table[ lower + 8]  := 37.06;
			IQ_Table[ lower + 9]  := 127.06;
			IQ_Table[ lower + 10]  := 58.24;
			IQ_Table[ lower + 11]  := 148.24;
			IQ_Table[ lower + 12]  := 10.59;
			IQ_Table[ lower + 13]  := 105.88;
			IQ_Table[ lower + 14]  := 42.35;
			IQ_Table[ lower + 15]  := 132.35;
			IQ_Table[ lower + 16]  := 26.47;
			IQ_Table[ lower + 17]  := 111.18;
			IQ_Table[ lower + 18]  := 52.94;
			IQ_Table[ lower + 19]  := 142.94;
			IQ_Table[ lower + 20]  := 5.29;
			IQ_Table[ lower + 21]  := 95.29;
			IQ_Table[ lower + 22]  := 63.53;
			IQ_Table[ lower + 23]  := 153.53;
			IQ_Table[ lower + 24]  := 31.76;
			IQ_Table[ lower + 25]  := 121.76;
			IQ_Table[ lower + 26]  := 79.41;
			IQ_Table[ lower + 27]  := 169.41;
			IQ_Table[ lower + 28]  := 15.88;
			IQ_Table[ lower + 29]  := 100.59;
			IQ_Table[ lower + 30]  := 174.71;
			IQ_Table[ lower + 31]  := 74.12;
			IQ_Table[ lower + 32]  := 164.12;
			IQ_Table[ lower + 33]  := 84.71;

		70:
			IQ_Table[ lower + 0]  := 0.00;
			IQ_Table[ lower + 1]  := 92.57;
			IQ_Table[ lower + 2]  := 46.29;
			IQ_Table[ lower + 3]  := 133.71;
			IQ_Table[ lower + 4]  := 25.71;
			IQ_Table[ lower + 5]  := 113.14;
			IQ_Table[ lower + 6]  := 72.00;
			IQ_Table[ lower + 7]  := 159.43;
			IQ_Table[ lower + 8]  := 36.00;
			IQ_Table[ lower + 9]  := 123.43;
			IQ_Table[ lower + 10]  := 82.29;
			IQ_Table[ lower + 11]  := 169.71;
			IQ_Table[ lower + 12]  := 10.29;
			IQ_Table[ lower + 13]  := 102.86;
			IQ_Table[ lower + 14]  := 56.57;
			IQ_Table[ lower + 15]  := 144.00;
			IQ_Table[ lower + 16]  := 30.86;
			IQ_Table[ lower + 17]  := 118.29;
			IQ_Table[ lower + 18]  := 61.71;
			IQ_Table[ lower + 19]  := 149.14;
			IQ_Table[ lower + 20]  := 5.14;
			IQ_Table[ lower + 21]  := 97.71;
			IQ_Table[ lower + 22]  := 51.43;
			IQ_Table[ lower + 23]  := 154.29;
			IQ_Table[ lower + 24]  := 20.57;
			IQ_Table[ lower + 25]  := 108.00;
			IQ_Table[ lower + 26]  := 41.14;
			IQ_Table[ lower + 27]  := 128.57;
			IQ_Table[ lower + 28]  := 77.14;
			IQ_Table[ lower + 29]  := 164.57;
			IQ_Table[ lower + 30]  := 15.43;
			IQ_Table[ lower + 31]  := 138.86;
			IQ_Table[ lower + 32]  := 87.43;
			IQ_Table[ lower + 33]  := 174.86;
			IQ_Table[ lower + 34]  := 66.86;
		ELSE
			Calc_RoundCakeDivisionsTable := -1;
			RETURN;
	END_CASE
END_IF

IF g_bCurrentTableUniversal10 THEN
	IQ_Table[1] := IQ_Table[1] +5;
	IQ_Table[2] := IQ_Table[2] +5;
	IQ_Table[3] := IQ_Table[3] +5;
	IQ_Table[4] := IQ_Table[4] +5;
	IQ_Table[5] := IQ_Table[5] +5;
END_IF

Calc_RoundCakeDivisionsTable := I_Divisions / 2;
RETURN;

END_FUNCTION
